(* IEC 61131-3 sources: daoli-st-library/DL_Algo (part 11) *)

(* ---- FB_DL_DewpointReset.st ---- *)
//==============================================================================
// 功能块：FB_DL_DewpointReset ｜ 中文名称：依据室内露点重置冷冻水供水温度设定
// 所属子库：DL_Algo ｜ 版本：v1.0.0 ｜ 兼容：CODESYS V3.5+ / TwinCAT 3 / 汇川 InoProShop
// 功能描述：室内露点重置冷冻水供水温度设定：目标 = max(露点 + 安全余
//           量, 下限)，带上下限钳位与斜率限制（fRateKPerS，由
//           uDeltaTimeMs 显式积分，禁系统时间函数）。露点由
//           FC_DL_DewPointCalc 计算（Magnus-Tetens 常数唯一属主为
//           FC_DL_VaporPressureSat，R23 裁定）——只调用不复制。双出
//           口：结露风险（露点 + 余量超上限，供水被顶到上限，除湿能
//           力不足，如实外显不静默）与域外钳位提示。失能保持设定。
// 开源溯源 (Origin)：道莅 clean-room 防御性实现（仅借 OSCAT ROOM_CONTROL 行为定义/参数域，零代码行与符号名复制）
// 单位表：温度[摄氏度] / 相对湿度[%] / 余量[K] / 斜率[K每s] / 扫描间隔[ms]
// 错误码表：16#0002_3601 信息级（露点域外钳位：湿度钳 1~100、干球钳
//           −40~60、下游件域外提示，不置 bError）/ 16#0002_3602 信息
//           级（防结露下限生效，供水被顶到上限，除湿能力不足，不置
//           bError）/ 16#0002_3605 预留禁用（不得挪用）/ 16#0002_3610
//           故障级（供水上下限倒置或余量/斜率组态非法，置 bError）/
//           16#0002_3611 故障级（输入非有限或下游件数据不可信，置
//           bError）/ 16#0002_3612 预留禁用（不得挪用）
// 状态机：E_DL_DewpointResetState（eIdle=0 / eTrack=10 / eCondRisk=20 /
//           eFault=99），CASE 含 ELSE 兜底，ELSE 复用 3611（§3 未为本
//           件单列兜底槽，不得越段加码）并回上限安全侧
// 边界行为：① 湿度钳 1~100、干球钳 −40~60（下游件承诺域），钳位发生
//           → 信息 3601；② 露点 + 余量大于供水上限 → bCondRisk :=
//           TRUE + 信息 3602，设定被顶到上限（如实反映「制冷量再低
//           也压不住露点」，不静默），退出条件两条：风险消失回追踪相
//           或失能回待机；③ fChwMinC 大于等于 fChwMaxC 或余量小于 0
//           或斜率非正 → 故障 3610；④ 非有限（NaN 自反判 + Inf 幅值
//           上限判，R79）→ 故障 3611，设定回供水上限安全侧（防结露
//           优先，冷却失效由上位温控回路告警，不静默）；⑤ 下游露点
//           件 uErrorId 非零或 bInRange 为假（预钳位后正常不可达，防
//           御路径）→ 复用信息 3601 且露点取干球温度保守估计（热力学
//           事实：露点不超过干球），下游信息级不升格（R115 纪律反向
//           适用：信息安全侧不得放大）；⑥ 失能 → 保持设定 + bValid :=
//           FALSE（供水温度突变会导致除湿振荡）；⑦ 斜率限制用
//           uDeltaTimeMs 显式积分，间隔为 0 本拍不动；⑧ 首拍设定从
//           下限起坡（首拍不出未知值）。
// 修订历史：v1.0.0 2026-11-17 首版（R25 派单 · §4.9）
//==============================================================================
(*------------------------------------------------------------------------------
 * 枚举: E_DL_DewpointResetState（归属 DL_Algo，与 FB_DL_DewpointReset 同文件）
 *----------------------------------------------------------------------------*)
TYPE E_DL_DewpointResetState :
(
    eIdle     := 0,   // 失能/待机：设定保持 / Idle: setpoint held
    eTrack    := 10,  // 斜率追踪：向目标设定限速逼近 / Track: rate-limited approach to target
    eCondRisk := 20,  // 结露风险：目标超上限，供水顶上限 / Condensation risk: target above ceiling, supply pinned
    eFault    := 99   // 故障兜底态：组态非法/非有限/非法状态，设定回上限 / Fault fallback, setpoint at ceiling
);
END_TYPE
FUNCTION_BLOCK FB_DL_DewpointReset
VAR_INPUT
    fRoomTempC    : LREAL;                     // 室内干球温度 [摄氏度] / Room dry-bulb temperature [degC]
    fRoomRhPct    : LREAL;                     // 室内相对湿度 [百分数] / Room relative humidity [percent]
    fChwMinC      : LREAL := 7.0;              // 供水设定下限 [摄氏度] / Chilled-water setpoint floor [degC]
    fChwMaxC      : LREAL := 18.0;             // 供水设定上限 [摄氏度] / Chilled-water setpoint ceiling [degC]
    fDewMarginK   : LREAL := 1.5;              // 防结露安全余量 [K] / Anti-condensation margin [K]
    fRateKPerS    : LREAL := 0.05;             // 设定斜率 [K每s] / Setpoint rate limit [K per s]
    uDeltaTimeMs  : UDINT;                     // 扫描间隔 [ms]，调用方注入，禁用系统时间函数 / Scan interval [ms], caller-injected
    bEnable       : BOOL;                      // 总使能 / Master enable
    bReset        : BOOL;                      // 复位，上升沿清状态与设定 / Reset, rising edge clears state and setpoint
END_VAR
VAR_OUTPUT
    fChwSetC      : LREAL;                     // 冷冻水供水温度设定 [摄氏度] / Chilled-water supply setpoint [degC]
    fDewPointC    : LREAL;                     // 室内露点 [摄氏度]，下游件计算透传 / Room dew point [degC], passed through
    fMarginK      : LREAL;                     // 当前供水设定相对露点裕量 [K] / Margin of setpoint over dew point [K]
    bCondRisk     : BOOL;                      // 露点超出可调范围，除湿能力不足 / Dew point beyond adjustable range, dehumidification short
    bAtMin        : BOOL;                      // 设定贴下限 / Setpoint at floor
    bAtMax        : BOOL;                      // 设定贴上限 / Setpoint at ceiling
    eErr          : UDINT;                     // 错误码，0 = 无错，码位 16#0002_3601 起信息级、16#0002_3610 起故障级（分带见错误码表） / Error code, 0 = no error, band info/fault per the code table
    bError        : BOOL;                      // 故障级标志，仅故障级错误置位 / Fault-class flag, set only on fault-level codes
    bValid        : BOOL;                      // 设定数据可用标志，失能/故障闸显式 FALSE / Setpoint usable flag, explicit FALSE on disable/fault gates
    eState        : E_DL_DewpointResetState;   // 主状态机当前状态 / Current state of the main state machine
END_VAR
VAR
    fbReset       : R_TRIG;                    // 复位上升沿检测实例 / Reset rising edge detector
    fRhClamped    : LREAL;                     // 钳位后湿度 [百分数] / Clamped humidity [percent]
    fTempClamped  : LREAL;                     // 钳位后干球 [摄氏度] / Clamped dry-bulb [degC]
    bDomainClamp  : BOOL;                      // 本拍发生域外钳位 / Domain clamp occurred this scan
    fTempReal     : REAL;                      // 干球降精度暂存 [摄氏度] / Dry-bulb staging in REAL precision
    fRhReal       : REAL;                      // 湿度降精度暂存 [百分数] / Humidity staging in REAL precision
    fDewReal      : REAL;                      // 露点返回值暂存 [摄氏度] / Dew-point return staging in REAL precision
    uDewErr       : UDINT;                     // 下游件错误码暂存 / Downstream error code staging
    fVaporPa      : REAL;                      // 下游件水汽压暂存 [Pa]（诊断透传）/ Downstream vapor pressure staging [Pa]
    bDewInRange   : BOOL;                      // 下游件域内标志暂存 / Downstream in-domain flag staging
    bDewOk        : BOOL;                      // 下游件结果可用判据 / Downstream result usable predicate
    fTargetC      : LREAL;                     // 钳位前目标设定 [摄氏度] / Pre-limit target setpoint [degC]
    fStepK        : LREAL;                     // 本拍允许步长 [K] / Allowed step this scan [K]
    fDeltaK       : LREAL;                     // 本拍目标增量 [K] / Target delta this scan [K]
    fDeltaApplied : LREAL;                     // 本拍实际增量 [K]（步长限幅后）/ Applied delta after rate limit [K]
    bFirstScan    : BOOL := TRUE;              // 首拍初始化标志 / First-scan initialization flag
END_VAR
VAR CONSTANT
    DL_DPR_CODE_INFO_1 : UDINT := 16#0002_3601;   // 信息级槽 1（露点域外钳位） / info slot 1
    DL_DPR_CODE_INFO_2 : UDINT := 16#0002_3602;   // 信息级槽 2（防结露下限生效） / info slot 2
    DL_DPR_CODE_RSV_1  : UDINT := 16#0002_3605;   // 预留禁用（不得挪用） / reserved, do not use
    DL_DPR_CODE_FLT_1  : UDINT := 16#0002_3610;   // 故障级槽 1（供水界倒置或组态非法） / fault slot 1
    DL_DPR_CODE_FLT_2  : UDINT := 16#0002_3611;   // 故障级槽 2（输入非有限） / fault slot 2
    DL_DPR_CODE_RSV_2  : UDINT := 16#0002_3612;   // 预留禁用（不得挪用） / reserved, do not use
    DL_DP_ZERO    : LREAL := 0.0;              // 零值常量，避免裸字面量 [—] / Zero constant, avoids a bare literal
    DL_DP_TOL     : LREAL := 1.0E-6;           // 浮点比较容差 [—] / Float comparison tolerance
    DL_DP_INF     : LREAL := 1.7976931348623157E308;  // LREAL 幅值上限，Inf 判据 / LREAL magnitude ceiling, Inf criterion
    DL_DP_RH_MIN  : LREAL := 1.0;              // 湿度钳位下限 [百分数] / Humidity clamp floor [percent]
    DL_DP_RH_MAX  : LREAL := 100.0;            // 湿度钳位上限 [百分数] / Humidity clamp ceiling [percent]
    DL_DP_T_MIN   : LREAL := -40.0;            // 干球钳位下限 [摄氏度]，下游件承诺域 / Dry-bulb clamp floor, downstream promised domain
    DL_DP_T_MAX   : LREAL := 60.0;             // 干球钳位上限 [摄氏度] / Dry-bulb clamp ceiling [degC]
    DL_DP_MS_PER_S : LREAL := 1000.0;          // 毫秒转秒系数 [s/ms] / Ms-to-s factor
END_VAR

(*------------------------------------------------------------------------------
 * 段 1｜无条件刷新区（红线 5）：复位沿检测在任何分支之外周期调用
 *----------------------------------------------------------------------------*)
fbReset(CLK := bReset);                        // 复位沿检测无条件刷新 / reset edge refreshed unconditionally

(*------------------------------------------------------------------------------
 * 段 2｜复位沿处理（改写置于沿后，防吞沿 R39）
 *----------------------------------------------------------------------------*)
IF fbReset.Q THEN
    eState  := E_DL_DewpointResetState.eIdle;
    eErr    := 16#0000_0000;                   // 复位清码 / reset clears code
    bError  := FALSE;                          // 复位清故障 / reset clears fault
    bCondRisk := FALSE;                        // 结露风险标志清 / condensation risk cleared
    bAtMin  := FALSE;                          // 贴下限清 / at-floor cleared
    bAtMax  := FALSE;                          // 贴上限清 / at-ceiling cleared
    bFirstScan := TRUE;                        // 重新首拍化 / re-initialize first scan
    fChwSetC := DL_DP_ZERO;                    // 设定清零待首拍初始化 / setpoint zeroed, awaits first-scan init
END_IF

(*------------------------------------------------------------------------------
 * 段 3｜非有限输入闸（浮点引脚逐个：NaN 自反判 + Inf 幅值上限判，R79）
 *       命中即设定回上限安全侧（防结露优先）
 *----------------------------------------------------------------------------*)
IF (fRoomTempC <> fRoomTempC) OR (ABS(fRoomTempC) >= DL_DP_INF)
   OR (fRoomRhPct <> fRoomRhPct) OR (ABS(fRoomRhPct) >= DL_DP_INF)
   OR (fChwMinC <> fChwMinC) OR (ABS(fChwMinC) >= DL_DP_INF)
   OR (fChwMaxC <> fChwMaxC) OR (ABS(fChwMaxC) >= DL_DP_INF)
   OR (fDewMarginK <> fDewMarginK) OR (ABS(fDewMarginK) >= DL_DP_INF)
   OR (fRateKPerS <> fRateKPerS) OR (ABS(fRateKPerS) >= DL_DP_INF) THEN
    eState  := E_DL_DewpointResetState.eFault;
    eErr    := DL_DPR_CODE_FLT_2;              // 故障级：输入非有限 / fault: non-finite input
    bError  := TRUE;                           // 故障级必置 bError（R45 配对）/ fault-class pairs with bError
    bValid  := FALSE;                          // 输出不可用 / outputs unusable
    fChwSetC := fChwMaxC;                      // 设定回上限安全侧（防结露优先）/ setpoint to ceiling, safe side
    bCondRisk := FALSE;                        // 故障态不判结露风险 / risk not judged in fault
    bAtMin := FALSE;                           // 贴限撤 / at-floor withdrawn
    bAtMax := TRUE;                            // 贴上限如实外显 / at-ceiling shown truthfully
    fDewPointC := DL_DP_ZERO;                  // 露点出口清零 / dew-point output zeroed
    fMarginK := DL_DP_ZERO;                    // 裕量出口清零 / margin output zeroed
    RETURN;
END_IF

(*------------------------------------------------------------------------------
 * 段 4｜组态合法性闸（供水界倒置/余量小于 0/斜率非正）
 *----------------------------------------------------------------------------*)
IF (fChwMinC >= fChwMaxC) OR (fDewMarginK < DL_DP_ZERO) OR (fRateKPerS <= DL_DP_TOL) THEN
    eState  := E_DL_DewpointResetState.eFault;
    eErr    := DL_DPR_CODE_FLT_1;              // 故障级：供水上下限倒置或组态非法 / fault: band inverted or config invalid
    bError  := TRUE;                           // 故障级必置 bError（R45 配对）/ fault-class pairs with bError
    bValid  := FALSE;                          // 输出不可用 / outputs unusable
    fChwSetC := fChwMaxC;                      // 设定回上限安全侧（防结露优先）/ setpoint to ceiling, safe side
    bCondRisk := FALSE;                        // 故障态不判结露风险 / risk not judged in fault
    bAtMin := FALSE;                           // 贴限撤 / at-floor withdrawn
    bAtMax := TRUE;                            // 贴上限如实外显 / at-ceiling shown truthfully
    fDewPointC := DL_DP_ZERO;                  // 露点出口清零 / dew-point output zeroed
    fMarginK := DL_DP_ZERO;                    // 裕量出口清零 / margin output zeroed
    RETURN;
END_IF

(*------------------------------------------------------------------------------
 * 段 5｜首拍初始化：设定从下限起坡（首拍不出未知值）
 *----------------------------------------------------------------------------*)
IF bFirstScan THEN
    fChwSetC := fChwMinC;                      // 首拍设定 = 下限 / first-scan setpoint = floor
    bFirstScan := FALSE;                       // 初始化完成 / initialization done
END_IF

(*------------------------------------------------------------------------------
 * 段 6｜域钳位（湿度 1~100、干球 −40~60，下游件承诺域）+ 露点组合调用
 *       （FC_DL_DewPointCalc，每拍恰好一次，只调用不复制）
 *----------------------------------------------------------------------------*)
fRhClamped := fRoomRhPct;                      // 湿度工作副本 / humidity working copy
fTempClamped := fRoomTempC;                    // 干球工作副本 / dry-bulb working copy
bDomainClamp := FALSE;                         // 钳位标志逐拍重判 / clamp flag re-judged per scan
IF fRhClamped < DL_DP_RH_MIN THEN
    fRhClamped := DL_DP_RH_MIN;                // 湿度钳下限 / humidity clamped to floor
    bDomainClamp := TRUE;                      // 钳位发生 / clamped
END_IF
IF fRhClamped > DL_DP_RH_MAX THEN
    fRhClamped := DL_DP_RH_MAX;                // 湿度钳上限 / humidity clamped to ceiling
    bDomainClamp := TRUE;                      // 钳位发生 / clamped
END_IF
IF fTempClamped < DL_DP_T_MIN THEN
    fTempClamped := DL_DP_T_MIN;               // 干球钳下限 / dry-bulb clamped to floor
    bDomainClamp := TRUE;                      // 钳位发生 / clamped
END_IF
IF fTempClamped > DL_DP_T_MAX THEN
    fTempClamped := DL_DP_T_MAX;               // 干球钳上限 / dry-bulb clamped to ceiling
    bDomainClamp := TRUE;                      // 钳位发生 / clamped
END_IF
fTempReal := LREAL_TO_REAL(fTempClamped);      // 干球降精度显式转换 / dry-bulb explicit narrowing
fRhReal := LREAL_TO_REAL(fRhClamped);          // 湿度降精度显式转换 / humidity explicit narrowing
fDewReal := FC_DL_DewPointCalc(fTempC := fTempReal, fRhPct := fRhReal,
                               uErrorId => uDewErr, fVaporPa => fVaporPa,
                               bInRange => bDewInRange);  // 露点组合调用，返回值即露点 [摄氏度] / dew-point call, return is the dew point
bDewOk := (uDewErr = 16#0000_0000) AND bDewInRange;    // 下游可用判据 / downstream usable predicate
IF bDewOk THEN
    fDewPointC := fDewReal;                    // 露点出口透传 / dew-point output pass-through
ELSE
    fDewPointC := fTempClamped;                // 防御路径：露点取干球保守估计（露点不超过干球）/ defensive: dry-bulb conservative estimate
    bDomainClamp := TRUE;                      // 下游域外提示并入钳位信息（不升格）/ downstream hint merged into clamp info
END_IF

(*------------------------------------------------------------------------------
 * 段 7｜目标计算：max(露点 + 余量, 下限)，超上限则顶上限并置结露风险
 *----------------------------------------------------------------------------*)
fTargetC := fDewPointC + fDewMarginK;          // 防结露目标 = 露点 + 余量 [摄氏度] / target = dew point plus margin
IF fTargetC < fChwMinC THEN
    fTargetC := fChwMinC;                      // 低于下限抬到下限 / below floor raised to floor
END_IF
IF fTargetC > fChwMaxC THEN
    fTargetC := fChwMaxC;                      // 超上限顶到上限 / above ceiling pinned to ceiling
END_IF

(*------------------------------------------------------------------------------
 * 段 8｜状态机：CASE 含 ELSE 兜底（非法状态 → 复用 3611 + 回上限，安全侧）
 *----------------------------------------------------------------------------*)
CASE eState OF

    E_DL_DewpointResetState.eIdle:
        bValid := FALSE;                       // 失能闸显式不可用（R72）/ explicit FALSE on disable gate
        bCondRisk := FALSE;                    // 待机不判风险 / risk not judged in idle
        bAtMin := FALSE;                       // 贴限撤 / at-floor withdrawn
        bAtMax := FALSE;                       // 贴限撤 / at-ceiling withdrawn
        eErr := 16#0000_0000;                  // 待机无错 / no error in idle
        bError := FALSE;                       // 待机无故障 / no fault in idle
        IF bEnable THEN
            eState := E_DL_DewpointResetState.eTrack;  // 使能进追踪相 / enable enters track
        END_IF

    E_DL_DewpointResetState.eTrack:
        bValid := TRUE;                        // 追踪相设定可用 / setpoint usable in track
        eErr := 16#0000_0000;                  // 追踪相先清码 / track clears code first
        bError := FALSE;                       // 追踪相先清故障 / track clears fault first
        IF bDomainClamp THEN
            eErr := DL_DPR_CODE_INFO_1;        // 信息级：露点域外钳位 / info: dew-point domain clamp
        END_IF
        IF NOT bEnable THEN
            eState := E_DL_DewpointResetState.eIdle;   // 失能回待机（设定保持）/ disable returns to idle, setpoint held
            bValid := FALSE;                   // 失能闸显式不可用 / explicit FALSE on disable gate
        ELSE
            fStepK := fRateKPerS * UDINT_TO_LREAL(uDeltaTimeMs) / DL_DP_MS_PER_S;  // 本拍步长 = 斜率乘时长 [K]，间隔 0 即不动 / step = rate times interval
            fDeltaK := fTargetC - fChwSetC;    // 目标增量 [K] / target delta [K]
            IF ABS(fDeltaK) <= fStepK THEN
                fDeltaApplied := fDeltaK;      // 一步到位 / single-step arrival
            ELSIF fDeltaK > DL_DP_ZERO THEN
                fDeltaApplied := fStepK;       // 正向限速 / positive rate-limited
            ELSE
                fDeltaApplied := -fStepK;      // 反向限速 / negative rate-limited
            END_IF
            fChwSetC := fChwSetC + fDeltaApplied;      // 限速逼近目标 / rate-limited approach
            bAtMin := ABS(fChwSetC - fChwMinC) < DL_DP_TOL;    // 贴下限（容差比较）/ at-floor with tolerance
            bAtMax := ABS(fChwSetC - fChwMaxC) < DL_DP_TOL;    // 贴上限（容差比较）/ at-ceiling with tolerance
            IF (fDewPointC + fDewMarginK) > fChwMaxC + DL_DP_TOL THEN
                eState := E_DL_DewpointResetState.eCondRisk;   // 露点超上限转结露风险相 / dew point beyond ceiling enters risk
            END_IF
        END_IF

    E_DL_DewpointResetState.eCondRisk:
        bValid := TRUE;                        // 风险相设定可用（顶上限值）/ setpoint usable in risk (pinned value)
        fChwSetC := fChwMaxC;                  // 供水被顶到上限（除湿能力不足，如实外显）/ supply pinned to ceiling
        bCondRisk := TRUE;                     // 结露风险标志 / condensation risk flag
        bAtMin := FALSE;                       // 贴下限撤 / at-floor withdrawn
        bAtMax := TRUE;                        // 贴上限如实外显 / at-ceiling shown truthfully
        eErr := DL_DPR_CODE_INFO_2;            // 信息级：防结露下限生效 / info: anti-condensation limit active
        bError := FALSE;                       // 信息级不置 bError / info never raises bError
        IF NOT bEnable THEN
            eState := E_DL_DewpointResetState.eIdle;   // 失能回待机（第二条退出条件）/ disable returns to idle, second exit
            bValid := FALSE;                   // 失能闸显式不可用 / explicit FALSE on disable gate
            bCondRisk := FALSE;                // 风险标志清 / risk flag cleared
        ELSIF (fDewPointC + fDewMarginK) <= fChwMaxC + DL_DP_TOL THEN
            eState := E_DL_DewpointResetState.eTrack;  // 风险消失回追踪相（第一条退出条件）/ risk gone, first exit to track
        END_IF

    ELSE
        eState := E_DL_DewpointResetState.eFault;  // 非法状态兜底 / illegal-state fallback
        eErr := DL_DPR_CODE_FLT_2;             // 兜底复用故障级槽 2（§3 未单列兜底槽，不得越段加码）/ fallback reuses fault slot 2
        bError := TRUE;                        // 故障级必置 bError / fault-class pairs with bError
        bValid := FALSE;                       // 输出不可用 / outputs unusable
        fChwSetC := fChwMaxC;                  // 设定回上限安全侧（防结露优先）/ setpoint to ceiling, safe side
        bCondRisk := FALSE;                    // 风险标志清 / risk flag cleared
        bAtMin := FALSE;                       // 贴限撤 / at-floor withdrawn
        bAtMax := TRUE;                        // 贴上限如实外显 / at-ceiling shown truthfully
END_CASE

(*------------------------------------------------------------------------------
 * 段 9｜裕量出口：当前供水设定相对露点裕量 [K]（负值即结露，可观测）
 *----------------------------------------------------------------------------*)
fMarginK := fChwSetC - fDewPointC;             // 裕量 = 设定 − 露点 [K] / margin = setpoint minus dew point
END_FUNCTION_BLOCK

(* ---- FB_DL_Differentiator.st ---- *)
(*==============================================================================
 * 组件名称 (Component)  : FB_DL_Differentiator
 * 所属子库 (Sublibrary) : DL_Algo
 * 当前版本 (Version)    : 1.0.1
 * 兼容性   (Platform)   : CODESYS 3.5 / TwinCAT 3 / 汇川 InoProShop / Machine Expert
 *                         仅依赖 Standard.library（LIMIT / MIN / MAX / ABS），零厂商方言
 * 功能描述 (Function)   : 带一阶低通滤波的实用微分器：差分商 (fIn - fInPrev)/fDt
 *                         计算变化率，后接一阶低通抑制高频噪声放大（纯差分对
 *                         采样噪声增益 1/fDt，会放大毛刺）。输出变化率限幅
 *                         （rRateMin/rRateMax）防异常尖峰误触发趋势报警。
 *                         现场用途：温度变化速率监控（趋势报警前级）、压装
 *                         速度计算、液位升降速率。
 * 开源溯源 (Origin)     : 原创实现。组合语义对应西门子 LGF 的差分商块与
 *                         PT1 滤波器串联的公开行为定义，clean-room 编写，
 *                         未复制任何厂商私有库源码。
 * 本文件内含       : TYPE  E_DL_DiffState（配套枚举，归属 DL_Algo）
 *                    FB    FB_DL_Differentiator
 * 依赖     (Depends)    : 无 DL_ 内部依赖；Standard.library: LIMIT / MIN / MAX / ABS
 * 红线自检 (Redline)    : R1 ✓ 零全局变量表与外部变量引用 ｜ R2 ✓ 零物理 IO 地址直写
 *                         R3 ✓ 纯 IEC 61131-3 ｜ R4 ✓ 防除零+钳位+非有限值拒绝
 *                         R5 ✓ 全变量中英双语同行注释 ｜ R6 ✓ 四态 ENUM+CASE+ELSE
 *                         R7 N/A（无定时器/边沿实例）
 * 【边界披露 / Boundary disclosure】
 *   B1 除零防御：fDt 走公共钳位（<10ms 钳位 10ms 置 16#0002_0002），恒大于零。
 *   B2 tFiltTime 超上限 60s：钳位并置 16#0002_1401；tFiltTime=0 为合法直通
 *      （输出原始差分商，不置故障）。
 *   B3 rRateMin > rRateMax：自动对调并置 16#0002_0001。
 *   B4 输入非有限值：本拍拒绝、清历史（bHistValid=FALSE）、输出归零，置
 *      16#0002_0004；下一有效拍重新同步端点，绝不输出伪造速率。
 *   B5 首扫同步 fInPrev := fIn、输出 0，防上电尖峰。
 *   B6 低通系数 fAlpha 显式钳位 0..1；fTfEff + fDt 恒 > 0（分母安全）。
 * 【验收向量 / Acceptance vectors】
 *   V1  fIn 每拍 +1.0（tSampleTime=100MS，即 10 EU/s 恒速）→ fRawRate=10 EU/s，
 *       fRateOut 数拍内收敛到 10 EU/s、bValid=TRUE
 *   V2  fIn 阶跃 +50 一拍 → fRawRate=500 EU/s 单拍尖峰，fRateOut 按
 *       tFiltTime=500MS 平滑，峰值明显低于 500（噪声抑制效果）
 *   V3  fIn 恒定 → fRateOut 收敛到 0
 *   V4  rRateMax=20，V1 → fRateOut 钳位 20 EU/s
 *   V5  tFiltTime=0 → fRateOut=fRawRate（直通，无故障码）
 *   V6  tFiltTime=65S → 钳位 60S、16#0002_1401
 *   V7  fIn=NaN → 16#0002_0004，fRateOut=0、bValid=FALSE
 * 修订历史 (Revision)   :
 *   2026-11-15  v1.0.0  首版入库（Round 04 · Phase 3 · DL_Algo 批次）
 *   2026-11-15  v1.0.1  阶段五终审精修：首扫初始化标志判据修复（原判据恒假
 *                       为死代码），首扫同步端点改为显式可审计路径
 *============================================================================*)

(*-----------------------------------------------------------------------------
 * 枚举: E_DL_DiffState（归属 DL_Algo，与 FB_DL_Differentiator 同文件）
 * 含义: 微分器状态机离散状态。数值步长留空位便于后续插态而不破坏已有工程。
 *----------------------------------------------------------------------------*)
TYPE E_DL_DiffState :
(
    eInit  := 0,   // 初始化态：首扫或失历史，同步端点、输出清零 / Init state, sync endpoint, output zero
    eRun   := 10,  // 运行态：差分商 + 低通滤波逐拍计算 / Run state, difference quotient with low-pass per scan
    eTrack := 20,  // 跟踪态：输出立即跟随 fTrackValue / Track state, output follows track value instantly
    eFault := 99   // 故障兜底态：非法状态拦截，自动回初始化 / Fault fallback, auto recover to init
);
END_TYPE

(*==============================================================================
 * 功能块: FB_DL_Differentiator
 * 调用约定: 每个扫描周期无条件调用一次；bTrack 使能时输出立即跟随 fTrackValue。
 * 无状态泄漏: 全部状态驻留于实例私有 VAR，可多实例并行互不影响。
 * 噪声披露: 输出滞后 ≈ tFiltTime；tFiltTime 越小噪声抑制越弱，建议
 *           tFiltTime >= 5 × 采样周期（本块默认 500ms @ 100ms 采样）。
 *============================================================================*)
FUNCTION_BLOCK FB_DL_Differentiator
VAR_INPUT
    bEnable     : BOOL := FALSE;      // 使能标志，FALSE 时输出 0 / Enable flag, FALSE forces output to zero
    fIn         : REAL := 0.0;        // 被微分量 [EU]，如温度/位置/液位 / Differentiated input [EU]
    tFiltTime   : TIME := T#500MS;    // 速率低通时间常数 [s]，0 = 原始差分直通 / Rate low-pass time constant [s], 0 = raw pass
    rRateMin    : REAL := -1.0E10;    // 速率下限 [EU/s]，大于上限时自动对调 / Rate lower limit [EU/s], swapped if greater
    rRateMax    : REAL := 1.0E10;     // 速率上限 [EU/s]，小于下限时自动对调 / Rate upper limit [EU/s], swapped if smaller
    bTrack      : BOOL := FALSE;      // 跟踪使能，TRUE 时输出立即跟随 fTrackValue / Track enable, output follows track value
    fTrackValue : REAL := 0.0;        // 跟踪值 [EU/s]，投切无扰动基准 / Track value [EU/s], bumpless transfer reference
    tSampleTime : TIME := T#100MS;    // 采样周期 [s]，小于 10ms 钳位为 10ms / Sample time [s], clamped to 10ms
END_VAR
VAR_OUTPUT
    fRateOut    : REAL;               // 变化率输出 [EU/s]，滤波并限幅 / Rate output [EU/s], filtered and limited
    fRawRate    : REAL;               // 未滤波原始速率 [EU/s]，诊断 / Raw unfiltered rate [EU/s] for diagnostics
    bValid      : BOOL;               // 输出有效标志（端点已同步且有真实差分）/ Output valid flag
    bError      : BOOL;               // 故障标志（瞬时，逐拍重算） / Fault flag, transient, recomputed every scan
    uErrorId    : UDINT;              // 故障码，0 = 无故障 / Error code, 0 = no error
END_VAR
VAR
    fInPrev     : REAL;               // 上一拍被微分量 [EU]，差分端点 / Previous input [EU], difference endpoint
    fTfEff      : REAL;               // 钳位后滤波时间常数 [s] / Clamped filter time constant [s]
    fAlpha      : REAL;               // 低通滤波系数 [0..1] / Low-pass filter coefficient [0..1]
    fDt         : REAL;               // 折算后的采样周期 [s] / Converted sample period [s]
    bInFinite   : BOOL;               // 本拍输入有限值标志 / Input finite validity flag this scan
    bHistValid  : BOOL;               // 端点历史有效标志 / Endpoint history valid flag
    bInit       : BOOL;               // 首扫标志 / First scan flag
    eState      : E_DL_DiffState;     // 主状态机当前状态 / Current state of the main state machine
END_VAR
VAR CONSTANT
    DL_DIFF_TF_MAX : REAL := 60.0;    // 滤波时间常数上限 [s] / Filter time constant upper limit [s]
    DL_DIFF_EPS    : REAL := 1.0E-6;  // 分母安全容差 / Denominator safety tolerance
END_VAR

(*------------------------------------------------------------------------------
 * 段 1｜公共参数处理（通用约定 0-1/0-2/0-3）：周期钳位、滤波常数钳位、量程对调
 *      Common handling: sample time clamp, filter constant clamp, limit swap
 *-----------------------------------------------------------------------------*)
uErrorId := 16#0000_0000;               // 故障码逐拍重算 / Error code recomputed every scan
bError   := FALSE;                      // 故障标志逐拍重算 / Fault flag recomputed every scan

IF tSampleTime < T#10MS THEN
    fDt      := TIME_TO_REAL(T#10MS) / 1000.0; // 非法周期钳位为 10ms（边界 B1 防除零）/ Illegal period clamped to 10ms
    uErrorId := 16#0002_0002;           // 采样周期非法已钳位 / Sample time illegal, clamped
ELSE
    fDt      := TIME_TO_REAL(tSampleTime) / 1000.0; // 周期换算为秒 [s] / Period converted to seconds [s]
END_IF

fTfEff := TIME_TO_REAL(tFiltTime) / 1000.0; // 滤波常数换算为秒 [s] / Filter constant converted to seconds [s]
IF fTfEff < 0.0 THEN
    fTfEff   := 0.0;                    // 负值钳位为直通 / Negative clamped to pass-through
    uErrorId := 16#0002_1401;           // 滤波时间常数非法已钳位 / Filter time constant illegal, clamped
END_IF
IF fTfEff > DL_DIFF_TF_MAX THEN
    fTfEff   := DL_DIFF_TF_MAX;         // 超上限钳位（边界 B2）/ Over-limit clamped
    uErrorId := 16#0002_1401;           // 滤波时间常数非法已钳位 / Filter time constant illegal, clamped
END_IF

IF rRateMin > rRateMax THEN
    rRateMin := rRateMin + rRateMax;    // 三步对调第一步：求和 / Swap step one: sum
    rRateMax := rRateMin - rRateMax;    // 三步对调第二步：得旧下限 / Swap step two: old lower limit
    rRateMin := rRateMin - rRateMax;    // 三步对调第三步：得旧上限 / Swap step three: old upper limit
    uErrorId := 16#0002_0001;           // 参数越界已对调 / Limits out of order, swapped
END_IF

(*------------------------------------------------------------------------------
 * 段 2｜输入合法性（边界 B4）：非有限值拒绝并清历史，输出归零防伪造速率
 *      Input validity: non-finite rejected, history cleared, output zeroed
 *-----------------------------------------------------------------------------*)
bInFinite := NOT (fIn <> fIn) AND (ABS(fIn) <= 1.0E30); // NaN 判别 + 幅值防御 / NaN check plus magnitude guard

IF NOT bInFinite THEN
    uErrorId   := 16#0002_0004;         // 输入非有限值已拒绝 / Non-finite input rejected
    bHistValid := FALSE;                // 清历史端点 / Clear endpoint history
    fRateOut   := 0.0;                  // 输出归零 / Output zeroed
    fRawRate   := 0.0;                  // 原始速率归零 / Raw rate zeroed
    bValid     := FALSE;                // 有效标志清零 / Valid flag cleared
    eState     := eInit;                // 回初始化态重新同步 / Back to init for re-sync
END_IF

(*------------------------------------------------------------------------------
 * 段 3｜跟踪与首扫（约定 0-6）：端点同步、输出归零，防上电尖峰（边界 B5）
 *      Tracking and first scan: endpoint synced, output zeroed against power-up spike
 *-----------------------------------------------------------------------------*)
IF NOT bInit THEN
    IF bInFinite THEN
        fInPrev := fIn;                 // 端点同步当前输入 / Endpoint synced to current input
        bHistValid := TRUE;             // 历史有效 / History valid
    END_IF
    fRateOut := 0.0;                    // 输出清零 / Output zeroed
    fRawRate := 0.0;                    // 原始速率清零 / Raw rate zeroed
    bValid   := FALSE;                  // 首扫无真实差分 / No real difference on first scan
    eState   := eInit;                  // 回初始化态 / Back to init state
    bInit    := TRUE;                   // 首扫标志置位 / First scan flag set
END_IF

IF bTrack THEN
    fRateOut := LIMIT(rRateMin, fTrackValue, rRateMax); // 输出立即跟随跟踪值并限幅 / Output follows track value with limits
    IF bInFinite THEN
        fInPrev := fIn;                 // 端点同步当前输入 / Endpoint synced to current input
    END_IF
    bHistValid := TRUE;                 // 历史有效 / History valid
    bValid     := TRUE;                 // 跟踪输出视为有效 / Tracked output considered valid
    eState     := eTrack;               // 跟踪态 / Track state
END_IF

(*------------------------------------------------------------------------------
 * 段 4｜使能失效语义：输出归零、清历史，恢复后从初始化态重新同步
 *      Disabled semantics: output zeroed, history cleared, re-sync after enable
 *-----------------------------------------------------------------------------*)
IF NOT bEnable THEN
    fRateOut   := 0.0;                  // 输出归零 / Output zeroed
    fRawRate   := 0.0;                  // 原始速率归零 / Raw rate zeroed
    bValid     := FALSE;                // 有效标志清零 / Valid flag cleared
    bHistValid := FALSE;                // 清历史端点 / Clear endpoint history
    eState     := eInit;                // 回初始化态 / Back to init state
ELSE
    (*--------------------------------------------------------------------------
     * 段 5｜主状态机（红线 R6）：四态 ENUM + CASE + ELSE 兜底
     *     Main state machine: four-state ENUM + CASE with mandatory ELSE fallback
     *-------------------------------------------------------------------------*)
    CASE eState OF

        eInit:  // 初始化态：端点同步、输出 0，下拍进入运行态（边界 B5）/ Init: sync endpoint, output zero
            IF bInFinite THEN
                fInPrev := fIn;             // 端点同步当前输入 / Endpoint synced to current input
                bHistValid := TRUE;         // 历史有效 / History valid
            END_IF
            fRateOut := 0.0;                // 输出清零 / Output zeroed
            fRawRate := 0.0;                // 原始速率清零 / Raw rate zeroed
            bValid   := FALSE;              // 本拍无真实差分 / No real difference this scan
            eState   := eRun;               // 进入运行态 / Enter run state

        eRun:  // 运行态：差分商 + 低通滤波（边界 B1 分母安全）/ Run: difference quotient with low-pass
            IF NOT bHistValid THEN
                fInPrev := fIn;             // 历史失效先重建端点 / Rebuild endpoint when history invalid
                bHistValid := TRUE;         // 历史恢复有效 / History restored
                fRateOut := 0.0;            // 输出先归零防尖峰 / Output zeroed against spike
                fRawRate := 0.0;            // 原始速率归零 / Raw rate zeroed
            ELSE
                fRawRate := (fIn - fInPrev) / fDt; // 原始差分商 [EU/s] / Raw difference quotient [EU/s]
                IF fTfEff <= DL_DIFF_EPS THEN
                    fAlpha := 1.0;          // 零滤波常数直通（边界 B2 合法）/ Zero constant pass-through
                ELSE
                    fAlpha := fDt / (fTfEff + fDt); // 一阶低通系数 [0..1] / First-order low-pass coefficient
                    fAlpha := MIN(MAX(fAlpha, 0.0), 1.0); // 系数显式钳位（边界 B6）/ Coefficient explicitly clamped
                END_IF
                fRateOut := fRateOut + fAlpha * (fRawRate - fRateOut); // 低通递推 [EU/s] / Low-pass recursion [EU/s]
                fRateOut := LIMIT(rRateMin, fRateOut, rRateMax); // 速率限幅 / Rate limited
                fInPrev  := fIn;            // 端点更新 / Endpoint updated
                bValid   := TRUE;           // 输出有效 / Output valid
            END_IF

        eTrack:  // 跟踪态：输出已由段 3 跟随，释放后回运行态 / Track: output follows, resume run after release
            IF NOT bTrack THEN
                eState := eRun;             // 释放跟踪，恢复计算 / Tracking released, resume computing
            END_IF

        eFault:  // 故障兜底态：输出归零并回初始化态（无锁死）/ Fault fallback: output zeroed, recover to init
            fRateOut := 0.0;                // 输出归零 / Output zeroed
            eState   := eInit;              // 自动恢复初始化 / Auto recover to init

        ELSE  // 非法状态拦截：任何未定义状态一律进故障态并置码 / Illegal state interception
            eState   := eFault;             // 强制故障态 / Force fault state
            uErrorId := 16#0002_0005;       // 非法状态兜底 / Illegal state fallback
            bError   := TRUE;               // 故障标志置位 / Fault flag set

    END_CASE;
END_IF
END_FUNCTION_BLOCK

(* ---- FB_DL_DisturbanceObserver.st ---- *)
(*
  FB_DL_DisturbanceObserver  —  模型法负载扰动观测器 / Model-based load disturbance observer
  分类 Category : DL_Algo
  码位 Code     : 16#02_3_81
  版本 Version  : 1.0.0
  来源标签 Tag  : t2-4-s7-motion
  溯源 Source   : S7 Motion Control 语义借鉴 · clean-room 实现，仅借分类/参数域/命名，未复制源码行
  功能 Function : 1) 标称模型逆（J·dω/dt ÷ Kt）折算等效电流，与指令电流之差乘 Kt 得扰动转矩估计；
                  2) 估计量经一阶 Q 滤波（委托 FB_DL_LowPassFilter）去噪后输出；
                  3) 补偿量按 fCompGain 加权并限幅到 ±fCompLimit，饱和置 bSaturated。
  边界 Boundary : ① fInertia / fTorqueConst / fQFilterTau / fRatedCurrentA 任一 <= 0 判组态错置码且不投运（防除零）；
                  ② 速度为零并持续超冻结窗 tZeroSpeedHold（本件常量 200 ms）时冻结估计（静止段无可观测加速度，防噪声灌入）；
                  ③ bEnable 下降沿清估计值与微分状态（R28-1 解除式 = bEnable 上升沿 + bReset，两路径均在引脚可满足）；
                  ④ 补偿限幅 fCompLimit 由引脚给出，不在本件硬编码；
                  ⑤ bEnable = FALSE 语义：输出降级为安全值 0 + 保持状态 eIdle，不冻结末值（R191 显式声明）。
  依赖 Depends  : FB_DL_LowPassFilter × 1（Q 滤波，每拍无条件调用）
  同拍双窗配比  : 冻结窗 tZeroSpeedHold = 200 ms 与 Q 滤波时间常数 fQFilterTau 同源于 fSampleDt；
                  配比约束 fQFilterTau <= 0.5 × tZeroSpeedHold 保证静止冻结前滤波器已收敛（R100）

  码表 Error codes（本件格 02_3_81，子码步进 +0x10）:
    16#0002_0281 故障级：组态非法（惯量 / 转矩常数 / 滤波时间常数 / 额定电流 <= 0，或采样周期 <= 0，或组态量非有限）
    16#0002_0291 故障级：相 ID 越界（枚举兜底路径，复用组态码段之外的单列码）
    16#0002_02A1 信息级：速度为零冻结估计 / 输入非有限本拍不更新（不置 bError）

  修订历史 Revision :
    2026-11-18  v1.0.0  R36 首版入库
*)

TYPE E_DL_ObserverState :
(
    eIdle  := 0,   // 空闲（未使能，输出降级为 0）/ Idle, outputs degraded to zero
    eRun   := 10,  // 观测运行 / Observer running
    eHold  := 20,  // 静止冻结（速度为零超冻结窗）/ Frozen at zero speed
    eFault := 90   // 组态故障锁定（需 bReset 沿解除）/ Configuration fault locked
);
END_TYPE

FUNCTION_BLOCK FB_DL_DisturbanceObserver
VAR_INPUT
    bEnable        : BOOL := FALSE;              // 总使能，FALSE 时输出降级为 0 并回 eIdle / Master enable
    bReset         : BOOL := FALSE;              // 复位，上升沿清组态故障锁存 / Reset, clears latched fault
    fCmdOut        : REAL := 0.0;                // 控制器输出（力矩指令）[% 额定力矩] / Controller output [% rated torque]
    fRatedCurrentA : REAL := 10.0;               // 额定电流 [A]，域 > 0 / Rated current [A], domain > 0
    fMeasSpeed     : REAL := 0.0;                // 实测转速 [rpm]，带符号 / Measured speed [rpm]
    fInertia       : REAL := 0.001;              // 折算惯量 [kg·m²]，域 > 0 / Reflected inertia [kg·m²]
    fTorqueConst   : REAL := 1.0;                // 转矩常数 [N·m/A]，域 > 0 / Torque constant [N·m/A]
    fQFilterTau    : REAL := 0.005;              // Q 滤波时间常数 [s]，域 > 0 / Q-filter time constant [s]
    tSampleTime    : TIME := T#10MS;             // 采样周期 [ms 口径]，域 > 0 / Sampling period
    fCompGain      : REAL := 1.0;                // 补偿加权系数 [1]，域 >= 0 / Compensation gain
    fCompLimitPct  : REAL := 20.0;               // 补偿限幅 [%]，域 > 0 / Compensation limit [%]
    fEps           : REAL := 1.0E-6;             // 浮点判零容差 [1] / Floating zero tolerance
END_VAR
VAR_OUTPUT
    fDistTorqueEst : REAL;                       // 扰动转矩估计 [N·m] / Estimated disturbance torque [N·m]
    fCompOut       : REAL;                       // 补偿量输出 [%]，限幅后 / Compensation output [%]
    bSaturated     : BOOL;                       // 补偿限幅饱和标志（单拍）/ Compensation saturated, single scan
    bFrozen        : BOOL;                       // 静止冻结标志 / Frozen at zero speed
    bValid         : BOOL;                       // 估计有效标志（单拍）/ Estimate valid, single scan
    bError         : BOOL;                       // 故障标志，派生自锁存 / Fault flag derived from latch
    uErrorId       : UDINT;                      // 事件码，0 = 无事件 / Event code, 0 = no event
    eStateOut      : E_DL_ObserverState;         // 状态出口，段尾单点映射 / State mapped at tail
END_VAR
VAR
    fbQFilter      : FB_DL_LowPassFilter;        // Q 滤波实例（每拍无条件调用）/ Q-filter instance
    tonZeroSpeed   : TON;                        // 零速持续时间窗（本件常量 200 ms）/ Zero-speed dwell timer
    rtEnable       : R_TRIG;                     // 使能上升沿 / Enable rising edge
    rtReset        : R_TRIG;                     // 复位上升沿 / Reset rising edge
    _eState        : E_DL_ObserverState := E_DL_ObserverState.eIdle;  // 内部状态机当前态 / Internal phase
    _uFault        : UDINT;                      // 故障码锁存（仅复位沿清除）/ Latched fault code
    _uInfo         : UDINT;                      // 信息码，每拍重算 / Information code, recomputed each scan
    _bFault        : BOOL;                       // 故障锁存位 / Latched fault bit
    fSpeedPrev     : REAL;                       // 上一拍转速快照 [rpm]（不参与预清零）/ Speed snapshot, kept
    fAccelRpmS     : REAL;                       // 转速微分 [rpm/s] / Speed derivative [rpm/s]
    fAccelRadS     : REAL;                       // 角加速度 [rad/s²] / Angular acceleration [rad/s²]
    fCurrentNomA   : REAL;                       // 标称模型逆等效电流 [A] / Nominal model inverse current [A]
    fCurrentCmdA   : REAL;                       // 指令折算电流 [A] / Command current [A]
    fTorqueDistNm  : REAL;                       // 含噪扰动转矩 [N·m] / Raw disturbance torque [N·m]
    fDtSec         : REAL;                       // 采样周期秒值 [s] / Sampling period in seconds
    bFirstScan     : BOOL := TRUE;               // 首扫标志（微分初值用）/ First-scan flag for derivative
    bZeroSpeed     : BOOL;                       // 零速判定中间量 / Zero-speed predicate
    bCfgBad        : BOOL;                       // 组态非法聚合标志 / Configuration invalid aggregate
END_VAR
VAR CONSTANT
    DL_T_ZERO_HOLD : TIME  := T#200MS;   // 零速冻结窗 [ms]，本件声明常量 / Zero-speed freeze window
    DL_RPM2RAD     : REAL  := 0.1047197551;  // rpm 转 rad/s [rad/(s·rpm)] / rpm to rad/s factor
    DL_EPS         : REAL  := 1.0E-6;    // 判零容差 [1] / Zero tolerance
END_VAR

(* —— 段 0：定时器与边缘检测无条件周期刷新（禁置于分支内） —— *)
rtEnable(CLK := bEnable);                                      // 使能上升沿（每拍必调）
rtReset(CLK := bReset);                                        // 复位上升沿（每拍必调）
bZeroSpeed := bEnable AND (ABS(fMeasSpeed) < DL_EPS);          // 零速判定，门控挂状态量
tonZeroSpeed(IN := bZeroSpeed, PT := DL_T_ZERO_HOLD);          // 零速驻留计时（输入非字面 TRUE，具备复位路径）

(* —— 段 1：单拍标志预清零（只清单拍量，快照与锁存不入清单） —— *)
bSaturated := FALSE;      // 单拍标志：限幅饱和
bValid     := FALSE;      // 单拍标志：估计有效
bFrozen    := FALSE;      // 单拍标志：静止冻结
bError     := FALSE;      // 单拍标志：故障出口（段 6 由锁存派生重写）
_uInfo     := 0;          // 信息码每拍重算
fDtSec     := TIME_TO_REAL(tSampleTime) / 1000.0;   // 采样周期秒值 [s]

(* —— 段 2：复位沿清故障锁存（R188 可达清除路径） —— *)
IF rtReset.Q THEN
    _bFault := FALSE;     // 复位沿清锁存位
    _uFault := 0;         // 复位沿清锁存码
END_IF

(* —— 段 3：组态域闸（覆盖全部参与换算的引脚，R151） —— *)
bCfgBad := FALSE;
IF (fInertia <> fInertia) OR (fInertia <= 0.0) THEN
    bCfgBad := TRUE;      // 惯量非有限或 <= 0
END_IF
IF (fTorqueConst <> fTorqueConst) OR (fTorqueConst <= 0.0) THEN
    bCfgBad := TRUE;      // 转矩常数非有限或 <= 0
END_IF
IF (fQFilterTau <> fQFilterTau) OR (fQFilterTau <= 0.0) THEN
    bCfgBad := TRUE;      // 滤波时间常数非有限或 <= 0
END_IF
IF (fRatedCurrentA <> fRatedCurrentA) OR (fRatedCurrentA <= 0.0) THEN
    bCfgBad := TRUE;      // 额定电流非有限或 <= 0
END_IF
IF (fCompLimitPct <> fCompLimitPct) OR (fCompLimitPct <= 0.0) THEN
    bCfgBad := TRUE;      // 补偿限幅非有限或 <= 0
END_IF
IF (fEps <> fEps) OR (fEps <= 0.0) THEN
    bCfgBad := TRUE;      // 判零容差非有限或 <= 0
END_IF
IF tSampleTime <= T#0MS THEN
    bCfgBad := TRUE;      // 采样周期 <= 0（微分除零前置）
END_IF
IF bCfgBad THEN
    _uFault := 16#0002_0281;                              // 故障级：组态非法
    _bFault := TRUE;                                      // 锁存位置位（复位沿可清）
    bError := TRUE;                                       // 故障标志置位（R45 配对）
    _eState := E_DL_ObserverState.eFault;                 // 状态机进故障相
END_IF

(* —— 段 4：观测内核（仅无故障且使能时执行） —— *)
IF (NOT _bFault) AND bEnable AND (fDtSec > 0.0) THEN
    fCurrentCmdA := fCmdOut / 100.0 * fRatedCurrentA;                    // 指令折算电流 [A]
    IF bFirstScan THEN
        fSpeedPrev := fMeasSpeed;                                        // 首扫微分初值，防冲击
        bFirstScan := FALSE;                                             // 首扫标志唯一置假点
    END_IF
    fAccelRpmS := (fMeasSpeed - fSpeedPrev) / fDtSec;                    // 转速微分 [rpm/s]
    fAccelRadS := fAccelRpmS * DL_RPM2RAD;                               // 角加速度 [rad/s²]
    fSpeedPrev := fMeasSpeed;                                            // 快照更新（末行，不预清零）
    fCurrentNomA := fInertia * fAccelRadS / fTorqueConst;                // 标称模型逆等效电流 [A]（Kt 已证 > 0）
    fTorqueDistNm := (fCurrentCmdA - fCurrentNomA) * fTorqueConst;       // 含噪扰动转矩 [N·m]
    IF tonZeroSpeed.Q THEN
        _eState := E_DL_ObserverState.eHold;                             // 静止冻结相
        bFrozen    := TRUE;                                                // 冻结标志（出口 bFrozen，VAR_OUTPUT）
        _uInfo := 16#0002_02A1;                                         // 信息级：速度为零冻结估计
    ELSE
        _eState := E_DL_ObserverState.eRun;                             // 观测运行相
        fbQFilter(bEnable := TRUE, fIn := fTorqueDistNm, tTimeConst := REAL_TO_TIME(fQFilterTau * 1000.0),
                  tSampleTime := tSampleTime);                          // Q 滤波实例调用（每拍必调，单点单次）
        IF fbQFilter.bError THEN
            _eState := E_DL_ObserverState.eHold;                        // 滤波故障降级为冻结（降级不抛故障，R191 已声明）
        END_IF
    END_IF
ELSE
    _eState := E_DL_ObserverState.eIdle;                                // 未使能：降级为安全值（R191 声明）
    fSpeedPrev := fMeasSpeed;                                           // 快照跟随，防再使能冲击
    bFirstScan := TRUE;                                                 // 复位首扫标志（再使能重新取值）
END_IF

(* —— 段 5：状态机兜底（非法枚举值回 eIdle 并置故障级码） —— *)
CASE _eState OF
E_DL_ObserverState.eIdle:
    fCompOut := 0.0;                     // 空闲：补偿量降级为 0
    fDistTorqueEst := 0.0;               // 空闲：估计值清零
E_DL_ObserverState.eRun:
    fDistTorqueEst := fbQFilter.fOut;    // 运行：输出滤波后扰动估计 [N·m]
    fCompOut := -fCompGain * fDistTorqueEst / fTorqueConst / fRatedCurrentA * 100.0;  // 补偿量 [%]（Kt、额定电流已证 > 0）
    IF fCompOut > fCompLimitPct THEN
        fCompOut := fCompLimitPct;       // 上行限幅
        bSaturated := TRUE;              // 饱和标志
    ELSIF fCompOut < -fCompLimitPct THEN
        fCompOut := -fCompLimitPct;      // 下行限幅
        bSaturated := TRUE;              // 饱和标志
    END_IF
    bValid := TRUE;                      // 本拍估计有效
E_DL_ObserverState.eHold:
    fDistTorqueEst := 0.0;               // 冻结：不出新估计（静止段无可观测加速度）
    fCompOut := 0.0;                     // 冻结：补偿量 0
E_DL_ObserverState.eFault:
    fDistTorqueEst := 0.0;               // 故障：输出安全值
    fCompOut := 0.0;                     // 故障：输出安全值
ELSE
    _uFault := 16#0002_0291;             // 故障级：相 ID 越界（枚举兜底）
    _bFault := TRUE;                     // 锁存位置位
    bError := TRUE;                      // 故障标志置位（R45 配对）
    _eState := E_DL_ObserverState.eFault;  // 强制回故障相
    fDistTorqueEst := 0.0;               // 兜底输出安全值
    fCompOut := 0.0;                     // 兜底输出安全值
END_CASE

(* —— 段 6：出口单点映射（名实同源，故障码由锁存回放） —— *)
eStateOut := _eState;                    // 状态出口
IF _bFault THEN
    uErrorId := _uFault;                 // 故障锁存码回放（不在故障相按当下输入重推）
ELSE
    uErrorId := _uInfo;                  // 信息码
END_IF
bError := _bFault;                       // 故障出口派生自锁存（非擦除式覆盖）

END_FUNCTION_BLOCK

(* ---- FB_DL_DryingOvenZone.st ---- *)
// =====================================================================
// FB_DL_DryingOvenZone.st
// 烘箱 8 温区串级控温（比例 + 风量前馈 + 速率限幅 + 独立超温联锁）
// Drying oven 8-zone cascade temperature control FB
// 码位: 16#0002_371F ~ 16#0002_3723 (本件独占 5 槽)
// 修改记录: R29 初版 (按 DISPATCH_R29 序 5)
// =====================================================================
FUNCTION_BLOCK FB_DL_DryingOvenZone
VAR_INPUT
    bEnable         : BOOL  := FALSE;   // 使能 / Enable
    bReset          : BOOL  := FALSE;   // 复位 / Reset
    abZoneEnable    : ARRAY[1..8] OF BOOL;      // 8 区独立使能 / Per-zone enable
    afPv_C          : ARRAY[1..8] OF REAL;      // 8 区实测温度 -20~300 ℃ / Zone PV [degC]
    afSp_C          : ARRAY[1..8] OF REAL;      // 8 区设定温度 0~250 ℃ / Zone SP [degC]
    afKp            : ARRAY[1..8] OF REAL;      // 8 区比例增益 0.1~20 %/K / Zone gain [%/K]
    fFanPct         : REAL  := 0.0;     // 循环风量 0~100 % / Fan duty [%]
    fKff            : REAL  := 0.0;     // 风量前馈系数 0~1 %/% / Fan feedforward [%/%]
    fOvertemp_C     : REAL  := 260.0;   // 超温阈值 50~300 ℃ / Overtemperature limit [degC]
    fRateMax_pct_s  : REAL  := 5.0;     // 输出速率上限 >0 %/s / Output slew limit [%/s]
    bFanRun         : BOOL  := FALSE;   // 风机运行反馈 / Fan running
    tCycle          : TIME  := T#100MS; // 周期 T#10MS~T#2S / Cycle [s]
END_VAR
VAR_OUTPUT
    afOut_pct       : ARRAY[1..8] OF REAL;      // 8 区加热输出 0~100 % / Heater output [%]
    bOvertemp       : BOOL;             // 任一区超温（锁存）/ Any zone overtemp, latched
    uOvertempZone   : USINT;            // 首个超温区号 0=无 / First overtemp zone, 0=none
    bReady          : BOOL;             // 全部区进入带内 / All zones in band
    eState          : E_DL_OvenState;   // 状态 / State
    eErr            : UDINT;            // 错误码 / Error code
END_VAR
VAR
    uIdx            : UDINT;            // 区循环下标 / Zone loop index
    uZi             : INT;              // 1..8 数组下标 / Array subscript 1..8
    uZj2            : INT;              // 清零循环第二下标 / Second subscript for zero loops
    fDevK           : REAL;             // 区偏差 K / Zone deviation [K]
    fSpSafe         : REAL;             // 处理后设定（≤0 按 1 ℃）/ Sanitized SP [degC]
    fOutRaw         : REAL;             // 计算原始输出 / Raw computed output [%]
    fStepMax        : REAL;             // 单拍步长 / Max step per cycle [%]
    fStep           : REAL;             // 本拍实际步长 / Actual step this cycle [%]
    tCycleS         : REAL;             // 周期秒值（钳 ≥0.01）/ Cycle in seconds, clamped [s]
    bAllEnabled     : BOOL;             // 是否存在使能区 / Any zone enabled
    bFanBad         : BOOL;             // 风量非有限标记 / Fan duty non-finite flag
    fFanPctSafe     : REAL;             // 处理后风量 / Sanitized fan duty [%]
    bAnyOver        : BOOL;             // 本拍超温探测 / Overtemp detected this cycle
    uFirstOver      : USINT;            // 本拍首个超温区 / First overtemp zone this cycle
    xFirstScan      : BOOL := TRUE;     // 首扫标记 / First-scan flag
END_VAR

// ---------------------------------------------------------------------
// 代码位表（本件独占，勿复用）:
//   16#0002_371F 信息 正常运行
//   16#0002_3720 故障 任一 afPv_C/afSp_C 非有限，或 tCycle 非法
//   16#0002_3721 故障 fOvertemp_C ≤ 0 / fRateMax_pct_s ≤ 0 / 任一 afKp ≤ 0（组态错）
//   16#0002_3722 信息 bFanRun=FALSE → 前馈禁用（fKff 项按 0 计），调节继续
//   16#0002_3723 故障 任一区 afPv_C ≥ fOvertemp_C → 全输出清零、锁存，解除=bReset 且全部 PV < 阈值-5K
// ---------------------------------------------------------------------

// ---- 周期转秒并钳下限 / Cycle to seconds with clamp ----
tCycleS := TIME_TO_REAL(tCycle) / 1000.0;   // 秒值 / Seconds [s]
IF tCycleS < 0.01 THEN
    tCycleS := 0.01;    // 钳 ≥0.01 s 防步长爆炸 / Clamp minimum 10 ms
END_IF

// ---- 单拍步长 / Max step per cycle ----
fStepMax := fRateMax_pct_s * tCycleS;       // %/s × s = % / Step per cycle [%]

// ---- 超温锁存解除路径（必须可达，R28）：bReset 且全部 PV < 阈值-5K 回差 / Reset path with 5K hysteresis ----
IF bOvertemp AND bReset THEN
    bAnyOver := FALSE;          // 回差判据累加器 / Hysteresis accumulator
    FOR uIdx := 1 TO 8 DO
        uZi := UDINT_TO_INT(uIdx);              // 下标转换 / Subscript conversion
        IF afPv_C[uZi] >= (fOvertemp_C - 5.0) THEN
            bAnyOver := TRUE;   // 仍有区未回落 5K / Zone not cooled by 5K
        END_IF
    END_FOR
    IF NOT bAnyOver THEN
        bOvertemp     := FALSE; // 解除锁存 / Release latch
        uOvertempZone := 0;     // 区号清零 / Clear zone number
        eState := E_DL_OvenState.eIdle; // 回空闲 / Back to idle
    END_IF
END_IF

// ---- 非有限与周期合法性闸（故障级）/ Finite and cycle validity gate ----
IF (tCycle = T#0MS) OR (tCycleS > 2.0)
   OR (fFanPct <> fFanPct) OR (ABS(fFanPct) >= 1.0E12)
   OR (fKff <> fKff) OR (ABS(fKff) >= 1.0E12)
   OR (fOvertemp_C <> fOvertemp_C) OR (ABS(fOvertemp_C) >= 1.0E12)
   OR (fRateMax_pct_s <> fRateMax_pct_s) OR (ABS(fRateMax_pct_s) >= 1.0E12) THEN
    bOvertemp     := FALSE;     // 清锁存避免卡死 / Clear latch to avoid deadlock
    uOvertempZone := 0;         // 区号清零 / Clear zone
    FOR uZi := 1 TO 8 DO
        afOut_pct[uZi] := 0.0;  // 全输出清零（安全侧）/ Zero all outputs
    END_FOR
    bReady := FALSE;            // 就绪失效 / Not ready
    eState := E_DL_OvenState.eFault;    // 故障态（本闸不锁存，可自动恢复）/ Fault state
    eErr   := 16#0002_3720;     // 故障码 / Fault code
    RETURN;                     // 本拍结束 / End of cycle
END_IF

// ---- 各区 PV/SP 非有限逐个判界（多 ARRAY 按各自上界逐个判）/ Per-zone finite check ----
FOR uZi := 1 TO 8 DO
    IF (afPv_C[uZi] <> afPv_C[uZi]) OR (ABS(afPv_C[uZi]) >= 1.0E12)
       OR (afSp_C[uZi] <> afSp_C[uZi]) OR (ABS(afSp_C[uZi]) >= 1.0E12) THEN
        FOR uZj2 := 1 TO 8 DO
            afOut_pct[uZj2] := 0.0;  // 全输出清零 / Zero all outputs
        END_FOR
        bReady := FALSE;        // 就绪失效 / Not ready
        eState := E_DL_OvenState.eFault;    // 故障态 / Fault state
        eErr   := 16#0002_3720; // 故障码 / Fault code
        RETURN;                 // 本拍结束 / End of cycle
    END_IF
END_FOR

// ---- 组态错闸 / Configuration fault gate ----
IF (fOvertemp_C <= 0.0) OR (fRateMax_pct_s <= 0.0) THEN
    FOR uZi := 1 TO 8 DO
        afOut_pct[uZi] := 0.0;  // 全输出清零 / Zero all outputs
    END_FOR
    bReady := FALSE;            // 就绪失效 / Not ready
    eState := E_DL_OvenState.eFault;    // 故障态 / Fault state
    eErr   := 16#0002_3721;     // 故障码 / Fault code
    RETURN;                     // 本拍结束 / End of cycle
END_IF
FOR uZi := 1 TO 8 DO
    IF afKp[uZi] <= 0.0 THEN
        FOR uZj2 := 1 TO 8 DO
            afOut_pct[uZj2] := 0.0;  // 全输出清零 / Zero all outputs
        END_FOR
        bReady := FALSE;        // 就绪失效 / Not ready
        eState := E_DL_OvenState.eFault;    // 故障态 / Fault state
        eErr   := 16#0002_3721; // 故障码 / Fault code
        RETURN;                 // 本拍结束 / End of cycle
    END_IF
END_FOR

// ---- 首扫初始化（R16 首扫纪律）/ First-scan initialization ----
IF xFirstScan THEN
    FOR uZi := 1 TO 8 DO
        afOut_pct[uZi] := 0.0;  // 输出从 0 起步 / Outputs start at zero
    END_FOR
    xFirstScan := FALSE;        // 清首扫标记 / Clear flag
END_IF

// ---- 使能撤销：全区输出清零回空闲 / Disable: zero outputs and idle ----
IF NOT bEnable THEN
    FOR uZi := 1 TO 8 DO
        afOut_pct[uZi] := 0.0;  // 全输出清零 / Zero all outputs
    END_FOR
    bReady := FALSE;            // 就绪失效 / Not ready
    eState := E_DL_OvenState.eIdle;     // 空闲态 / Idle state
    eErr   := 16#0002_371F;     // 信息级：空闲正常 / Info: idle normal
    RETURN;                     // 本拍结束 / End of cycle
END_IF

// ---- 使能区存在性检查：全关 → eIdle 输出全 0 / No enabled zone → idle ----
bAllEnabled := FALSE;           // 累加器复位 / Reset accumulator
FOR uZi := 1 TO 8 DO
    IF abZoneEnable[uZi] THEN
        bAllEnabled := TRUE;    // 至少一区使能 / At least one zone enabled
    END_IF
END_FOR
IF NOT bAllEnabled THEN
    FOR uZi := 1 TO 8 DO
        afOut_pct[uZi] := 0.0;  // 全输出清零 / Zero all outputs
    END_FOR
    bReady := FALSE;            // 就绪失效 / Not ready
    eState := E_DL_OvenState.eIdle;     // 空闲态 / Idle state
    eErr   := 16#0002_371F;     // 信息级：空闲正常 / Info: idle normal
    RETURN;                     // 本拍结束 / End of cycle
END_IF

// ---- 风量前馈有效性：bFanRun=FALSE → 前馈项按 0 计 / Feedforward disabled without fan ----
bFanBad := FALSE;               // 标记复位 / Reset flag
fFanPctSafe := fFanPct;         // 原值采用 / Adopt as-is
IF NOT bFanRun THEN
    fFanPctSafe := 0.0;         // 前馈禁用（不是零输出）/ FF disabled, control continues
END_IF

// ---- 超温探测（超温优先于调节）/ Overtemp detection has priority ----
bAnyOver   := FALSE;            // 探测复位 / Reset detection
uFirstOver := 0;                // 首区清零 / Clear first zone
FOR uZi := 1 TO 8 DO
    IF afPv_C[uZi] >= fOvertemp_C THEN
        bAnyOver := TRUE;       // 探测到超温 / Overtemp found
        IF uFirstOver = 0 THEN
            uFirstOver := INT_TO_USINT(uZi);    // 记录首区 / Record first zone
        END_IF
    END_IF
END_FOR

IF bAnyOver THEN
    // 超温路径：全输出清零 + 故障锁存，绝不边降温边加热 / Overtemp: zero all, latch fault
    FOR uZi := 1 TO 8 DO
        afOut_pct[uZi] := 0.0;  // 全输出清零（安全侧）/ Zero all outputs
    END_FOR
    bOvertemp     := TRUE;      // 锁存 / Latch
    uOvertempZone := uFirstOver;    // 记首区 / First zone
    bReady        := FALSE;     // 就绪失效 / Not ready
    eState        := E_DL_OvenState.eFault;     // 故障态 / Fault state
    eErr          := 16#0002_3723;      // 故障码 / Fault code
    RETURN;                     // 本拍结束 / End of cycle
END_IF

// ---- 正常调节路径（eRun）：逐区比例 + 前馈 + 速率限幅 / Normal control path ----
eState := E_DL_OvenState.eRun;      // 运行态 / Run state
bReady := TRUE;                     // 就绪假设成立，区带外再翻 false / Assume ready, clear per zone
FOR uZi := 1 TO 8 DO
    IF abZoneEnable[uZi] THEN
        // 设定 ≤0 按 1 ℃ 处理（防冻结工况斜率无穷）/ SP ≤0 treated as 1 degC
        IF afSp_C[uZi] <= 0.0 THEN
            fSpSafe := 1.0;     // 防斜率无穷 / Guard slope
        ELSE
            fSpSafe := afSp_C[uZi]; // 原值 / As-is
        END_IF
        fDevK := fSpSafe - afPv_C[uZi];     // 偏差 = SP - PV / Deviation [K]
        // 比例项 + 风量前馈项 / Proportional + fan feedforward term
        fOutRaw := afKp[uZi] * fDevK + fKff * fFanPctSafe;  // 原始输出 [%]
        // 前馈禁用信息级（bFanRun=FALSE 且 fKff>0 时提示）/ FF disabled info
        IF (NOT bFanRun) AND (fKff > 0.0) THEN
            eErr := 16#0002_3722;   // 信息级：前馈禁用 / Info: FF disabled
        END_IF
        // 输出限幅 0~100 % / Clamp 0..100
        IF fOutRaw < 0.0 THEN
            fOutRaw := 0.0;     // 下限 / Lower clamp
        ELSIF fOutRaw > 100.0 THEN
            fOutRaw := 100.0;   // 上限 / Upper clamp
        END_IF
        // 速率限幅（单拍增量 ≤ fStepMax）/ Slew limit per cycle
        fStep := fOutRaw - afOut_pct[uZi];  // 期望步长 / Desired step [%]
        IF fStep > fStepMax THEN
            fStep := fStepMax;      // 正向限速 / Positive slew
        ELSIF fStep < -fStepMax THEN
            fStep := -fStepMax;     // 负向限速 / Negative slew
        END_IF
        afOut_pct[uZi] := afOut_pct[uZi] + fStep;   // 采纳步长 / Adopt step
        // 带内判（±2 K 带容差）/ In-band check (±2 K tolerance)
        IF ABS(fSpSafe - afPv_C[uZi]) > 2.0 THEN
            bReady := FALSE;    // 区带外 → 就绪失效 / Zone out of band
        END_IF
    ELSE
        afOut_pct[uZi] := 0.0;  // 禁用区输出保持 0 / Disabled zone output zero
    END_IF
END_FOR

// 未在任何分支改写 eErr 时补正常码 / Default normal code if untouched
IF eErr <> 16#0002_3722 THEN
    eErr := 16#0002_371F;       // 信息级：正常运行 / Info: normal run
END_IF

END_FUNCTION_BLOCK

(* ---- FB_DL_DuctLeakRateEst.st ---- *)
(*
  FB_DL_DuctLeakRateEst  —  风管漏风率估算（流量差法 + 静压修正 + 分级判据） / Duct air-leakage rate estimation by flow difference with static-pressure correction and class grading
  分类 Category : DL_Algo
  版本 Version  : 1.0.0
  来源 Source   : t1-2-oscat-building — 楼宇风管验收算法族深化
  溯源 Origin   : 道莅 clean-room 实现；漏风率 = 100×(送风-回风)/送风 与静压线性修正为公开暖通测试算法，未复制任何源码行
  功能 Function : 1) 流量差法：_fLeakPct = 100 × (fSupplyM3h - fReturnM3h) / fSupplyM3h，
                  分母 <= 1.0E-6 判非法（除零前置守卫）；
                  2) 静压修正：_fCorrPct = (fStaticPa - fStaticRefPa) / 10.0 × fPressCorrPctPer10Pa，
                  修正后 _fLeakCorr = _fLeakPct - _fCorrPct（除数为常量 10.0）；
                  3) 向上取整到 0.1%：先实数上限兜底 → 截断 → 按余量进位（正好整除不 +1，
                  禁 TRUNC(x)+1 写法，R28-2）；
                  4) 分级：A/B/C 三档阈值判据，越 C 档为不合格（eReject）。
                  5) 本件只有故障码、无信息码（派单硬约束）。
  接口 Interface: 输入送/回风量、静压与参考静压、修正系数、三档阈值；输出漏风率/分级/码
  边界 Boundary : ① 组态闸：fSupplyM3h <= 1.0E-6、fPressCorrPctPer10Pa < 0.0、
                  fClassAPct < 0.0 或 fClassBPct <= fClassAPct 或 fClassCPct <= fClassBPct
                  → 0386 锁存；② 送/回风量或静压非有限（NaN 自反 + Inf 差值自减）→ 0386 锁存；
                  ③ 取整前实数上限兜底（2.147483E9 对应 DINT 可表上界），防 LREAL→DINT 溢出；
                  ④ 回风量大于送风量时漏风率为负，按死区归 0（-0.05% 容差带），不判故障；
                  ⑤ 零全局耦合：无 GVL / VAR_EXTERNAL / %I %Q %M 直接地址。
  依赖 Depends  : Standard.library（R_TRIG）
  码表 Error codes（Algo 段 0002，故障窗口 0386；本件无信息码）:
    16#0002_0386 故障级：漏风率估算故障总码（组态非法 / 风量或静压非有限 / 送风量为零导致除零），
                 锁存至 bReset 上升沿；归因见 eCause，不新增码位（派单硬约束单码）
  修订历史 Revision :
    2026-11-19  v1.0.0  R43 首版（批次 2 · 序号 10）
*)

TYPE E_DL_DlrState :
(
    eIdle  := 0,      // 未使能待估算 / Idle, waiting evaluation
    eRun   := 10,     // 估算运行中 / Evaluation active
    eFault := 90      // 故障锁存相 / Fault latched phase
);
END_TYPE

TYPE E_DL_DlrClass :
(
    eNone    := 0,    // 未分级 / Not graded
    eClassA  := 1,    // A 级（最严） / Class A, tightest
    eClassB  := 2,    // B 级 / Class B
    eClassC  := 3,    // C 级 / Class C
    eReject  := 4     // 不合格（越 C 档） / Rejected, beyond class C
);
END_TYPE

TYPE E_DL_DlrCause :
(
    eNone      := 0,  // 无故障成因 / No cause
    eCfgIllegal:= 1,  // 组态非法 / Illegal configuration
    eNonFinite := 2,  // 输入非有限 / Non-finite input
    eDivZero   := 3   // 送风量过小（除零风险） / Supply flow too small
);
END_TYPE

FUNCTION_BLOCK FB_DL_DuctLeakRateEst
VAR_INPUT
    fSupplyM3h        : REAL := 0.0;      // 送风量 [m³/h]，域 > 0 / Supply air flow
    fReturnM3h        : REAL := 0.0;      // 回风量 [m³/h] / Return air flow
    fStaticPa         : REAL := 0.0;      // 实测静压 [Pa] / Measured static pressure
    fStaticRefPa      : REAL := 0.0;      // 参考静压 [Pa] / Reference static pressure
    fPressCorrPctPer10Pa : REAL := 0.5;   // 每 10 Pa 修正百分比 [%/10Pa]，域 >= 0 / Correction per 10 Pa
    fClassAPct        : REAL := 1.0;      // A 级上限 [%] / Class A limit
    fClassBPct        : REAL := 3.0;      // B 级上限 [%] / Class B limit
    fClassCPct        : REAL := 6.0;      // C 级上限 [%] / Class C limit
    fNegDeadbandPct   : REAL := 0.05;     // 负值死区 [%]，域 >= 0 / Negative deadband
    bEnable           : BOOL := FALSE;    // 估算使能（电平）[-] / Evaluation enable
    bReset            : BOOL := FALSE;    // 复位命令，上升沿清故障 [-] / Reset edge
END_VAR
VAR_OUTPUT
    eState            : E_DL_DlrState;    // 状态出口，段 6 单点映射 / State outlet
    eClass            : E_DL_DlrClass;    // 分级出口 / Grading outlet
    eCause            : E_DL_DlrCause;    // 故障成因出口（R190） / Fault cause outlet
    fLeakPct          : REAL;             // 原始漏风率 [%] / Raw leakage rate
    fLeakCorrPct      : REAL;             // 静压修正后漏风率 [%] / Corrected leakage rate
    fLeakCeilPct      : REAL;             // 向上取整到 0.1% 的漏风率 [%] / Ceil to 0.1 %
    bError            : BOOL;             // 故障锁存标志 [-] / Fault latch flag
    nErrId            : UDINT;            // 故障码，0 = 无故障（本件无信息码） / Fault code only
END_VAR
VAR
    _eState           : E_DL_DlrState := E_DL_DlrState.eIdle;     // 内部相位（CASE 唯一写入目标） / Internal phase
    _eClass           : E_DL_DlrClass := E_DL_DlrClass.eNone;     // 分级槽（每拍重算） / Grading slot
    _eCause           : E_DL_DlrCause := E_DL_DlrCause.eNone;     // 故障成因锁存（锁存量） / Latched cause
    rtReset           : R_TRIG;           // 复位沿实例，每周期无条件调用 / Reset edge
    _fDiffM3h         : REAL;             // 送回风量差 [m³/h]（当拍量） / Flow difference
    _fCorrPct         : REAL;             // 静压修正量 [%]（当拍量） / Pressure correction
    _fScaled          : REAL;             // 取整中间量（×10 后） / Scaling intermediate
    _iScaled          : DINT;             // 截断后整数（×10） / Truncated integer
    _bNonFin          : BOOL;             // 输入非有限当拍量 [-] / Non-finite input
    _bDivRisk         : BOOL;             // 除零风险当拍量 [-] / Divide risk
    _bCfgBad          : BOOL;             // 组态非法当拍量 [-] / Config illegal
    _bFault           : BOOL;             // 故障锁存位（锁存量） / Latched fault bit
    _uFault           : UDINT;            // 故障码锁存（锁存量） / Latched fault code
END_VAR

(* —— 段 0：沿实例无条件周期刷新 + 当拍量判据 —— *)
_bNonFin := (fSupplyM3h <> fSupplyM3h) OR (fReturnM3h <> fReturnM3h) OR (fStaticPa <> fStaticPa)
         OR ((fSupplyM3h - fSupplyM3h) <> (fSupplyM3h - fSupplyM3h))
         OR ((fReturnM3h - fReturnM3h) <> (fReturnM3h - fReturnM3h))
         OR ((fStaticPa - fStaticPa) <> (fStaticPa - fStaticPa));            // NaN 自反 + Inf 差值自减 / NaN and Inf detection
_bDivRisk := fSupplyM3h <= 1.0E-6;                                           // 送风量过小（除零风险） / Divide risk
_bCfgBad := _bDivRisk OR (fPressCorrPctPer10Pa < 0.0) OR (fClassAPct < 0.0)
            OR (fClassBPct <= fClassAPct) OR (fClassCPct <= fClassBPct)
            OR (fNegDeadbandPct < 0.0);                                      // 组态非法当拍量 / Config illegal
rtReset(CLK := bReset);                                                      // 复位沿，每拍必调 / Reset edge

(* —— 段 1：单拍量预清零（锁存量不入清单；分级槽每拍重算） —— *)
eClass := E_DL_DlrClass.eNone;      // 分级出口缺省未分级 / Grading default
eCause := _eCause;                  // 成因出口映射（锁存量回放，段 6 复核） / Cause outlet
fLeakPct := 0.0;                    // 原始漏风率缺省 0 / Raw rate default
fLeakCorrPct := 0.0;                // 修正后漏风率缺省 0 / Corrected rate default
fLeakCeilPct := 0.0;                // 取整漏风率缺省 0 / Ceil rate default
nErrId := 16#0000_0000;             // 故障码缺省无故障 / Fault code default

(* —— 段 2：复位沿 + 组态域闸 —— *)
IF rtReset.Q THEN                              // rtReset.Q = 当拍量 / current scan
    _bFault := FALSE;                          // 清故障锁存位（锁存量） / Clear fault latch
    _uFault := 16#0000_0000;                   // 清故障锁存码（锁存量） / Clear fault code
    _eCause := E_DL_DlrCause.eNone;            // 清成因（锁存量） / Clear cause
    IF _eState = E_DL_DlrState.eFault THEN
        _eState := E_DL_DlrState.eIdle;        // 故障相迁出：回未使能 / Fault exit to idle
    END_IF
END_IF
IF _bNonFin THEN                               // 非有限锁存（独立归因） / Non-finite latch
    _uFault := 16#0002_0386;                   // 故障级：估算故障总码 / Algo fault code
    _eCause := E_DL_DlrCause.eNonFinite;       // 归因：非有限 / Cause: non-finite
    _bFault := TRUE;                           // 标志与码位配对（R45） / Flag paired with code
END_IF
IF _bCfgBad THEN                               // 组态域闸 / Config gate
    _uFault := 16#0002_0386;
    IF _bDivRisk THEN
        _eCause := E_DL_DlrCause.eDivZero;     // 归因：除零风险 / Cause: divide risk
    ELSE
        _eCause := E_DL_DlrCause.eCfgIllegal;  // 归因：组态非法 / Cause: illegal config
    END_IF
    _bFault := TRUE;
END_IF

(* —— 段 3：漏风率与分级（仅无故障时计算；除数为已校验正域） —— *)
IF (NOT _bFault) AND (_eState = E_DL_DlrState.eRun) THEN
    _fDiffM3h := fSupplyM3h - fReturnM3h;                          // 流量差 / Flow difference
    fLeakPct := 100.0 * _fDiffM3h / fSupplyM3h;                    // 原始漏风率（分母已守卫） / Raw rate
    _fCorrPct := (fStaticPa - fStaticRefPa) / 10.0 * fPressCorrPctPer10Pa;   // 静压修正（除常量 10.0） / Correction
    fLeakCorrPct := fLeakPct - _fCorrPct;                          // 修正后漏风率 / Corrected rate
    IF (fLeakCorrPct < 0.0) AND (ABS(fLeakCorrPct) <= fNegDeadbandPct) THEN
        fLeakCorrPct := 0.0;                                       // 负值死区归 0 / Negative deadband
    END_IF
    _fScaled := fLeakCorrPct * 10.0;                               // 放大 10 倍进入整数域 / Scale by ten
    IF _fScaled >= 2.147483E9 THEN                                 // 实数上限兜底（DINT 可表上界） / Real upper guard
        _fScaled := 2.147483E9;
    ELSIF _fScaled <= -2.147483E9 THEN                             // 实数下限兜底 / Real lower guard
        _fScaled := -2.147483E9;
    END_IF
    _iScaled := LREAL_TO_DINT(LREAL(_fScaled));                    // 截断取整 / Truncate
    IF LREAL(_iScaled) < LREAL(_fScaled) - 1.0E-9 THEN             // 余量进位（正好整除不进位） / Ceiling by remainder
        _iScaled := _iScaled + 1;
    END_IF
    fLeakCeilPct := DINT_TO_REAL(_iScaled) * 0.1;                  // 还原为 0.1% 步长 / Restore 0.1 % step
    IF fLeakCeilPct <= fClassAPct THEN
        _eClass := E_DL_DlrClass.eClassA;                          // A 级 / Class A
    ELSIF fLeakCeilPct <= fClassBPct THEN
        _eClass := E_DL_DlrClass.eClassB;                          // B 级 / Class B
    ELSIF fLeakCeilPct <= fClassCPct THEN
        _eClass := E_DL_DlrClass.eClassC;                          // C 级 / Class C
    ELSE
        _eClass := E_DL_DlrClass.eReject;                          // 不合格（ELSE 兜底） / Rejected fallback
    END_IF
END_IF

(* —— 段 4：故障解除式（R240；全当拍量）：rtReset.Q / NOT _bNonFin / NOT _bCfgBad —— *)
IF rtReset.Q AND (NOT _bNonFin) AND (NOT _bCfgBad) THEN
    _bFault := FALSE;                          // 清故障锁存位（锁存量） / Clear fault latch
    _uFault := 16#0000_0000;                   // 清故障锁存码（锁存量） / Clear fault code
    _eCause := E_DL_DlrCause.eNone;            // 清成因（锁存量） / Clear cause
END_IF

(* —— 段 4A：故障锁存相位迁移闸 —— *)
IF _bFault AND (_eState <> E_DL_DlrState.eFault) THEN
    _eState := E_DL_DlrState.eFault;           // 锁存即入故障相 / Latch enters fault phase
END_IF

(* —— 段 5：相位机（CASE 全覆盖 + ELSE 兜底） —— *)
CASE _eState OF

E_DL_DlrState.eIdle:
    IF bEnable AND (NOT _bFault) THEN          // 使能条件 / Enable gate
        _eState := E_DL_DlrState.eRun;         // 进估算相 / Enter evaluation
    END_IF

E_DL_DlrState.eRun:
    IF NOT bEnable THEN                        // 撤使能：回未使能（前置消失） / Disable returns idle
        _eState := E_DL_DlrState.eIdle;
    END_IF

E_DL_DlrState.eFault:
    ;                                          // 故障相：仅段 4 复位沿可迁出 / Only reset exits

ELSE
    _uFault := 16#0002_0386;                   // 故障级：非法相位兜底（归并总码） / Illegal phase fallback
    _eCause := E_DL_DlrCause.eCfgIllegal;      // 归因：相位非法归并组态 / Cause: phase illegal
    _bFault := TRUE;
    _eState := E_DL_DlrState.eFault;           // 强制回故障相 / Force fault phase

END_CASE

(* —— 段 6：出口单点映射（名实同源；锁存码回放，禁同拍抹除） —— *)
IF _bFault THEN
    nErrId := _uFault;                         // 故障锁存码回放 / Replay latched code
    eClass := E_DL_DlrClass.eNone;             // 故障相分级强制未分级 / Grading forced none
    fLeakCeilPct := 0.0;                       // 故障相取整值强制 0（安全侧） / Ceil forced zero
ELSE
    nErrId := 16#0000_0000;                    // 无故障：本件无信息码 / No fault, no info code
    eClass := _eClass;                         // 分级出口 / Grading outlet
END_IF
bError := _bFault;                             // 故障标志同源 / Flag from latch
eState := _eState;                             // 状态出口 / State outlet
eCause := _eCause;                             // 成因出口 / Cause outlet

END_FUNCTION_BLOCK

(* ---- FB_DL_DuctStaticReset.st ---- *)
//==============================================================================
// 功能块：FB_DL_DuctStaticReset ｜ 中文名称：风管静压设定重置
// 所属子库：DL_Algo ｜ 版本：v1.0.0 ｜ 兼容：CODESYS V3.5+ / TwinCAT 3 / 汇川 InoProShop
// 功能描述：风管静压设定重置（TSP 修剪侧单件）：最不利末端阀位落在目
//           标带 [100−band, 100) 视为合适（带内保持）；阀位顶满 100%
//           （超带）→ 设定按增益上抬；阀位低于带下沿 → 设定按增益下
//           调。设定变化经斜率限制（fRatePaPerS，由 uDeltaTimeMs 显式
//           积分，禁系统时间函数），上下限钳位。阀位反馈无效（bFbValid
//           为假）→ 保持上次设定并发 3502（信息级，不置 bError）；设
//           定已顶上限而阀位仍满开 → 3501 能力不足，不再继续抬设定。
//           只算设定值，不控变频器（风机调速由上位裁决，本件零执行输
//           出）。规格 §4.8 引脚表未给反馈有效性输入、但其边界行为③
//           与输出表均要求 bFbInvalid/3502 语义，故增补 VAR_INPUT
//           bFbValid（默认 TRUE）承载上游质量位（主动偏离披露，见修
//           订历史）。
// 开源溯源 (Origin)：道莅原创实现（参考 公开工程惯例 分类与参数域）
// 单位表：阀位[百分数] / 静压[Pa] / 目标带[百分数] / 增益[Pa每百分数] / 斜率[Pa每s] / 扫描间隔[ms]
// 错误码表：16#0002_3501 信息级（静压设定已顶上限且阀位仍全开，风机能
//           力不足，不再抬设定，不置 bError）/ 16#0002_3502 信息级（阀
//           位反馈无效，保持上次设定，不置 bError）/ 16#0002_3505 预留
//           禁用（不得挪用）/ 16#0002_3510 故障级（静压上下限倒置或
//           算法组态非法（带宽/增益/斜率非正），置 bError）/
//           16#0002_3511 故障级（输入非有限，置 bError，设定回下限安
//           全侧防过压）/ 16#0002_3512 预留禁用（不得挪用）
// 状态机：E_DL_DuctStaticState（eIdle=0 / eInBand=10 / eAdjustUp=20 /
//           eAdjustDown=30 / eFbHold=40 / eFault=99），CASE 含 ELSE 兜
//           底，ELSE 复用 3511（§3 未为本件单列兜底槽，不得越段加码）
//           并回下限安全侧
// 边界行为：① fStaticMinPa 大于等于 fStaticMaxPa 或带宽/增益/斜率非正
//           → 故障 3510；② 阀位域钳 0~100（轻域外按边界值照算）；
//           ③ 阀位反馈无效（bFbValid 为假）→ 保持上次设定 + 信息 3502，
//           挂 eFbHold 相，退出条件两条：反馈恢复（按带位回归工作相）
//           或失能（回待机）；④ 设定已达上限而阀位仍 100% → 信息 3501
//           + bAtLimit，不再继续抬设定；⑤ 斜率限制用 uDeltaTimeMs 显
//           式积分（LREAL 中间量，禁系统时间函数），uDeltaTimeMs 为 0
//           时本拍不动；⑥ 非有限（NaN 自反判 + Inf 幅值上限判，R79）
//           → 故障 3511，设定回 fStaticMinPa 安全侧（防过压）；⑦ 失
//           能 → 保持设定（静压突变会导致末端振荡）+ bValid := FALSE；
//           ⑧ 带语义披露：阀位落在 [100−band, 100) 带内保持，阀位 =
//           100% 视为顶带超限（需上抬），与验收向量 ①② 口径一致；
//           ⑨ 首拍设定从下限起坡（首拍不出未知值）。
// 修订历史：v1.0.0 2026-11-17 首版（R25 派单 · §4.8）
//==============================================================================
(*------------------------------------------------------------------------------
 * 枚举: E_DL_DuctStaticState（归属 DL_Algo，与 FB_DL_DuctStaticReset 同文件）
 *----------------------------------------------------------------------------*)
TYPE E_DL_DuctStaticState :
(
    eIdle       := 0,   // 失能/待机：设定保持，静压不突变 / Idle: setpoint held, no static jump
    eInBand     := 10,  // 阀位带内：设定保持 / In-band: damper within target band, setpoint held
    eAdjustUp   := 20,  // 阀位顶带：设定按斜率上抬 / Damper at band top: setpoint raised by rate
    eAdjustDown := 30,  // 阀位低于带：设定按斜率下调 / Damper below band: setpoint lowered by rate
    eFbHold     := 40,  // 反馈无效保持：设定保持，等反馈恢复 / Feedback-invalid hold: setpoint held
    eFault      := 99   // 故障兜底态：组态非法/非有限/非法状态，设定回下限 / Fault fallback, setpoint at floor
);
END_TYPE
FUNCTION_BLOCK FB_DL_DuctStaticReset
VAR_INPUT
    fWorstDamperPct : LREAL;                   // 最不利末端阀位 [百分数] / Worst-zone damper position [percent]
    fStaticMinPa  : LREAL;                     // 静压设定下限 [Pa] / Static setpoint floor [Pa]
    fStaticMaxPa  : LREAL;                     // 静压设定上限 [Pa] / Static setpoint ceiling [Pa]
    fBandPct      : LREAL := 10.0;             // 阀位目标带 [百分数]，带 = [100−band, 100) / Damper target band [percent]
    fGainPaPerPct : LREAL := 2.0;              // 增益 [Pa每百分数] / Gain [Pa per percent]
    fRatePaPerS   : LREAL := 5.0;              // 设定斜率 [Pa每s] / Setpoint rate limit [Pa per s]
    bFbValid      : BOOL := TRUE;              // 阀位反馈有效性质量位（规格补遗引脚，见修订历史）/ Damper feedback validity, spec-gap pin
    uDeltaTimeMs  : UDINT;                     // 扫描间隔 [ms]，调用方注入，禁用系统时间函数 / Scan interval [ms], caller-injected
    bEnable       : BOOL;                      // 总使能 / Master enable
    bReset        : BOOL;                      // 复位，上升沿清状态与设定 / Reset, rising edge clears state and setpoint
END_VAR
VAR_OUTPUT
    fStaticSetPa  : LREAL;                     // 静压设定 [Pa]，失能保持 / Static setpoint [Pa], held on disable
    bAtLimit      : BOOL;                      // 设定顶上限且阀位仍全开，能力不足 / Setpoint at ceiling with damper full open
    fErrPct       : LREAL;                     // 带偏差 [百分数]，阀位减带下沿，负 = 低于带 / Band deviation [percent], damper minus band floor
    bFbInvalid    : BOOL;                      // 阀位反馈无效标志 / Damper feedback invalid flag
    eErr          : UDINT;                     // 错误码，0 = 无错，码位 16#0002_3501 起信息级、16#0002_3510 起故障级（分带见错误码表） / Error code, 0 = no error, band info/fault per the code table
    bError        : BOOL;                      // 故障级标志，仅故障级错误置位 / Fault-class flag, set only on fault-level codes
    bValid        : BOOL;                      // 设定数据可用标志，失能/故障闸显式 FALSE / Setpoint usable flag, explicit FALSE on disable/fault gates
    eState        : E_DL_DuctStaticState;      // 主状态机当前状态 / Current state of the main state machine
END_VAR
VAR
    fbReset       : R_TRIG;                    // 复位上升沿检测实例 / Reset rising edge detector
    fDamperClamped : LREAL;                    // 钳位后阀位 [百分数] / Clamped damper position [percent]
    fBandFloor    : LREAL;                     // 带下沿 [百分数] / Band floor [percent]
    fStepPa       : LREAL;                     // 本拍允许步长 [Pa]（斜率乘时长）/ Allowed step this scan [Pa]
    fDeltaPa      : LREAL;                     // 本拍目标增量 [Pa]（增益乘带偏差）/ Target delta this scan [Pa]
    fDeltaApplied : LREAL;                     // 本拍实际增量 [Pa]（步长限幅后）/ Applied delta after rate limit [Pa]
    fSetTarget    : LREAL;                     // 限幅前目标设定 [Pa] / Pre-limit target setpoint [Pa]
    bFirstScan    : BOOL := TRUE;              // 首拍初始化标志 / First-scan initialization flag
END_VAR
VAR CONSTANT
    DL_DSR_CODE_INFO_1 : UDINT := 16#0002_3501;   // 信息级槽 1（顶上限且阀位全开） / info slot 1
    DL_DSR_CODE_INFO_2 : UDINT := 16#0002_3502;   // 信息级槽 2（反馈无效保持设定） / info slot 2
    DL_DSR_CODE_RSV_1  : UDINT := 16#0002_3505;   // 预留禁用（不得挪用） / reserved, do not use
    DL_DSR_CODE_FLT_1  : UDINT := 16#0002_3510;   // 故障级槽 1（静压界倒置或组态非法） / fault slot 1
    DL_DSR_CODE_FLT_2  : UDINT := 16#0002_3511;   // 故障级槽 2（输入非有限） / fault slot 2
    DL_DSR_CODE_RSV_2  : UDINT := 16#0002_3512;   // 预留禁用（不得挪用） / reserved, do not use
    DL_DS_ZERO    : LREAL := 0.0;              // 零值常量，避免裸字面量 [—] / Zero constant, avoids a bare literal
    DL_DS_TOL     : LREAL := 1.0E-6;           // 浮点比较容差 [—] / Float comparison tolerance
    DL_DS_INF     : LREAL := 1.7976931348623157E308;  // LREAL 幅值上限，Inf 判据 / LREAL magnitude ceiling, Inf criterion
    DL_DS_PCT_MAX : LREAL := 100.0;            // 阀位域上限 [百分数] / Damper domain ceiling [percent]
    DL_DS_MS_PER_S : LREAL := 1000.0;          // 毫秒转秒系数 [s/ms] / Ms-to-s factor
END_VAR

(*------------------------------------------------------------------------------
 * 段 1｜无条件刷新区（红线 5）：复位沿检测在任何分支之外周期调用
 *----------------------------------------------------------------------------*)
fbReset(CLK := bReset);                        // 复位沿检测无条件刷新 / reset edge refreshed unconditionally

(*------------------------------------------------------------------------------
 * 段 2｜复位沿处理（改写置于沿后，防吞沿 R39）
 *----------------------------------------------------------------------------*)
IF fbReset.Q THEN
    eState  := E_DL_DuctStaticState.eIdle;
    eErr    := 16#0000_0000;                   // 复位清码 / reset clears code
    bError  := FALSE;                          // 复位清故障 / reset clears fault
    bAtLimit := FALSE;                         // 贴限标志清 / at-limit flag cleared
    bFbInvalid := FALSE;                       // 反馈无效标志清 / invalid flag cleared
    bFirstScan := TRUE;                        // 重新首拍化 / re-initialize first scan
    fStaticSetPa := DL_DS_ZERO;                // 设定清零待首拍初始化 / setpoint zeroed, awaits first-scan init
END_IF

(*------------------------------------------------------------------------------
 * 段 3｜非有限输入闸（浮点引脚逐个：NaN 自反判 + Inf 幅值上限判，R79）
 *       命中即设定回下限安全侧（防过压）
 *----------------------------------------------------------------------------*)
IF (fWorstDamperPct <> fWorstDamperPct) OR (ABS(fWorstDamperPct) >= DL_DS_INF)
   OR (fStaticMinPa <> fStaticMinPa) OR (ABS(fStaticMinPa) >= DL_DS_INF)
   OR (fStaticMaxPa <> fStaticMaxPa) OR (ABS(fStaticMaxPa) >= DL_DS_INF)
   OR (fBandPct <> fBandPct) OR (ABS(fBandPct) >= DL_DS_INF)
   OR (fGainPaPerPct <> fGainPaPerPct) OR (ABS(fGainPaPerPct) >= DL_DS_INF)
   OR (fRatePaPerS <> fRatePaPerS) OR (ABS(fRatePaPerS) >= DL_DS_INF) THEN
    eState       := E_DL_DuctStaticState.eFault;
    eErr         := DL_DSR_CODE_FLT_2;             // 故障级：输入非有限 / fault: non-finite input
    bError       := TRUE;                      // 故障级必置 bError（R45 配对）/ fault-class pairs with bError
    bValid       := FALSE;                     // 输出不可用 / outputs unusable
    fStaticSetPa := fStaticMinPa;              // 设定回下限安全侧（防过压）/ setpoint to floor, safe side against overpressure
    bAtLimit := FALSE;                         // 故障态不判贴限 / at-limit not judged in fault
    bFbInvalid := FALSE;                       // 故障态不判反馈无效 / invalid not judged in fault
    fErrPct := DL_DS_ZERO;                     // 带偏差出口清零 / band deviation zeroed
    RETURN;
END_IF

(*------------------------------------------------------------------------------
 * 段 4｜组态合法性闸（静压界倒置/带宽/增益/斜率非正）
 *----------------------------------------------------------------------------*)
IF (fStaticMinPa >= fStaticMaxPa) OR (fBandPct <= DL_DS_TOL)
   OR (fGainPaPerPct <= DL_DS_TOL) OR (fRatePaPerS <= DL_DS_TOL) THEN
    eState       := E_DL_DuctStaticState.eFault;
    eErr         := DL_DSR_CODE_FLT_1;             // 故障级：静压上下限倒置或组态非法 / fault: static band inverted or config invalid
    bError       := TRUE;                      // 故障级必置 bError（R45 配对）/ fault-class pairs with bError
    bValid       := FALSE;                     // 输出不可用 / outputs unusable
    fStaticSetPa := fStaticMinPa;              // 设定回下限安全侧（防过压）/ setpoint to floor, safe side
    bAtLimit := FALSE;                         // 故障态不判贴限 / at-limit not judged in fault
    bFbInvalid := FALSE;                       // 故障态不判反馈无效 / invalid not judged in fault
    fErrPct := DL_DS_ZERO;                     // 带偏差出口清零 / band deviation zeroed
    RETURN;
END_IF

(*------------------------------------------------------------------------------
 * 段 5｜首拍初始化：设定从下限起坡（首拍不出未知值）
 *----------------------------------------------------------------------------*)
IF bFirstScan THEN
    fStaticSetPa := fStaticMinPa;              // 首拍设定 = 下限 / first-scan setpoint = floor
    bFirstScan := FALSE;                       // 初始化完成 / initialization done
END_IF

(*------------------------------------------------------------------------------
 * 段 6｜阀位钳位与带偏差计算（域钳 0~100，带下沿 = 100 − band）
 *----------------------------------------------------------------------------*)
fDamperClamped := fWorstDamperPct;             // 阀位工作副本 / working copy
IF fDamperClamped < DL_DS_ZERO THEN
    fDamperClamped := DL_DS_ZERO;              // 低于 0 钳入 / below zero clamped
END_IF
IF fDamperClamped > DL_DS_PCT_MAX THEN
    fDamperClamped := DL_DS_PCT_MAX;           // 高于 100 钳入 / above 100 clamped
END_IF
fBandFloor := DL_DS_PCT_MAX - fBandPct;        // 带下沿 = 100 − band [百分数] / band floor
fErrPct := fDamperClamped - fBandFloor;        // 带偏差：负 = 低于带，0~band = 带内，band = 顶带 / band deviation

(*------------------------------------------------------------------------------
 * 段 7｜状态机：CASE 含 ELSE 兜底（非法状态 → 复用 3511 + 回下限，安全侧）
 *----------------------------------------------------------------------------*)
CASE eState OF

    E_DL_DuctStaticState.eIdle:
        bValid := FALSE;                       // 失能闸显式不可用（R72）/ explicit FALSE on disable gate
        bAtLimit := FALSE;                     // 贴限标志清 / at-limit flag cleared
        bFbInvalid := FALSE;                   // 失能不判反馈无效 / invalid not judged in idle
        eErr := 16#0000_0000;                  // 待机无错 / no error in idle
        bError := FALSE;                       // 待机无故障 / no fault in idle
        IF bEnable THEN
            IF bFbValid THEN
                eState := E_DL_DuctStaticState.eInBand;        // 反馈有效进带内相 / valid feedback enters in-band
            ELSE
                eState := E_DL_DuctStaticState.eFbHold;        // 反馈无效进保持相 / invalid feedback enters hold
            END_IF
        END_IF

    E_DL_DuctStaticState.eInBand:
        bValid := TRUE;                        // 带内设定可用 / setpoint usable in band
        bAtLimit := FALSE;                     // 带内不判贴限 / at-limit not judged in band
        bFbInvalid := FALSE;                   // 反馈有效 / feedback valid
        eErr := 16#0000_0000;                  // 带内无错 / no error in band
        bError := FALSE;                       // 带内无故障 / no fault in band
        IF NOT bEnable THEN
            eState := E_DL_DuctStaticState.eIdle;      // 失能回待机（设定保持）/ disable returns to idle, setpoint held
            bValid := FALSE;                   // 失能闸显式不可用 / explicit FALSE on disable gate
        ELSIF NOT bFbValid THEN
            eState := E_DL_DuctStaticState.eFbHold;    // 反馈无效转保持相 / invalid feedback to hold phase
        ELSIF fErrPct >= fBandPct - DL_DS_TOL THEN     // 阀位顶满 100%（fErrPct 达 band 上沿即阀位 = 100）
            eState := E_DL_DuctStaticState.eAdjustUp;  // 顶带超限转上调相 / at band top enters adjust-up
        ELSIF fErrPct < -DL_DS_TOL THEN                // 阀位低于带下沿
            eState := E_DL_DuctStaticState.eAdjustDown;        // 低于带转下调相 / below band enters adjust-down
        END_IF

    E_DL_DuctStaticState.eAdjustUp:
        bValid := TRUE;                        // 上调相设定可用 / setpoint usable in adjust-up
        bFbInvalid := FALSE;                   // 反馈有效 / feedback valid
        IF NOT bEnable THEN
            eState := E_DL_DuctStaticState.eIdle;
            bValid := FALSE;                   // 失能闸显式不可用 / explicit FALSE on disable gate
        ELSIF NOT bFbValid THEN
            eState := E_DL_DuctStaticState.eFbHold;    // 反馈无效转保持相 / invalid feedback to hold phase
        ELSE
            fStepPa := fRatePaPerS * UDINT_TO_LREAL(uDeltaTimeMs) / DL_DS_MS_PER_S;  // 本拍步长 = 斜率乘时长 [Pa]，间隔 0 即不动 / step = rate times interval
            fDeltaPa := fGainPaPerPct * fErrPct;       // 目标增量 = 增益乘带偏差 [Pa] / target delta = gain times deviation
            IF fDeltaPa > fStepPa THEN
                fDeltaApplied := fStepPa;      // 斜率限幅 / rate-limited
            ELSE
                fDeltaApplied := fDeltaPa;     // 未触斜率 / within rate
            END_IF
            fSetTarget := fStaticSetPa + fDeltaApplied;        // 限幅前目标 [Pa] / pre-limit target
            IF fSetTarget >= fStaticMaxPa - DL_DS_TOL THEN
                fStaticSetPa := fStaticMaxPa;  // 钳到上限 / clamped to ceiling
                IF fDamperClamped >= DL_DS_PCT_MAX - DL_DS_TOL THEN
                    bAtLimit := TRUE;          // 设定顶上限且阀位仍全开：能力不足 / at ceiling with full-open damper
                    eErr := DL_DSR_CODE_INFO_1;        // 信息级：能力不足，不再抬设定 / info: capacity insufficient
                    bError := FALSE;           // 信息级不置 bError / info never raises bError
                ELSE
                    bAtLimit := FALSE;         // 阀位未满开，仅钳位 / damper not full, clamp only
                    eErr := 16#0000_0000;      // 清码 / clear code
                END_IF
            ELSE
                fStaticSetPa := fSetTarget;    // 未触上限照算 / below ceiling, apply
                bAtLimit := FALSE;             // 未贴限 / not at limit
                eErr := 16#0000_0000;          // 清码 / clear code
            END_IF
            IF fErrPct < fBandPct - DL_DS_TOL THEN     // 阀位离开顶带（需求消失退出）/ damper left band top
                IF fErrPct >= -DL_DS_TOL THEN
                    eState := E_DL_DuctStaticState.eInBand;    // 回带内相 / back to in-band
                ELSE
                    eState := E_DL_DuctStaticState.eAdjustDown;        // 落到带下方向 / fell below band
                END_IF
            END_IF
        END_IF

    E_DL_DuctStaticState.eAdjustDown:
        bValid := TRUE;                        // 下调相设定可用 / setpoint usable in adjust-down
        bAtLimit := FALSE;                     // 下调相不判贴限 / at-limit not judged in adjust-down
        bFbInvalid := FALSE;                   // 反馈有效 / feedback valid
        IF NOT bEnable THEN
            eState := E_DL_DuctStaticState.eIdle;
            bValid := FALSE;                   // 失能闸显式不可用 / explicit FALSE on disable gate
        ELSIF NOT bFbValid THEN
            eState := E_DL_DuctStaticState.eFbHold;    // 反馈无效转保持相 / invalid feedback to hold phase
        ELSE
            fStepPa := fRatePaPerS * UDINT_TO_LREAL(uDeltaTimeMs) / DL_DS_MS_PER_S;  // 本拍步长 [Pa] / step this scan
            fDeltaPa := fGainPaPerPct * (DL_DS_ZERO - fErrPct);        // 目标减量 = 增益乘带偏差绝对值 [Pa] / target decrement
            IF fDeltaPa > fStepPa THEN
                fDeltaApplied := fStepPa;      // 斜率限幅 / rate-limited
            ELSE
                fDeltaApplied := fDeltaPa;     // 未触斜率 / within rate
            END_IF
            fSetTarget := fStaticSetPa - fDeltaApplied;        // 限幅前目标 [Pa] / pre-limit target
            IF fSetTarget <= fStaticMinPa + DL_DS_TOL THEN
                fStaticSetPa := fStaticMinPa;  // 钳到下限 / clamped to floor
                eErr := 16#0000_0000;          // 清码 / clear code
            ELSE
                fStaticSetPa := fSetTarget;    // 未触下限照算 / above floor, apply
                eErr := 16#0000_0000;          // 清码 / clear code
            END_IF
            IF (fErrPct >= -DL_DS_TOL) AND (fErrPct < fBandPct - DL_DS_TOL) THEN
                eState := E_DL_DuctStaticState.eInBand;        // 回带相（需求消失退出）/ back to in-band when need gone
            END_IF
        END_IF

    E_DL_DuctStaticState.eFbHold:
        bValid := TRUE;                        // 保持相设定输出仍可用（保持值）/ usable in hold (held setpoint)
        bAtLimit := FALSE;                     // 保持相不判贴限 / at-limit not judged in hold
        bFbInvalid := TRUE;                    // 反馈无效标志保持 / invalid flag held
        eErr := DL_DSR_CODE_INFO_2;            // 信息级：反馈无效保持上次设定 / info: invalid feedback, setpoint held
        bError := FALSE;                       // 信息级不置 bError / info never raises bError
        IF NOT bEnable THEN
            eState := E_DL_DuctStaticState.eIdle;      // 失能回待机（第二条退出条件）/ disable returns to idle, second exit
            bValid := FALSE;                   // 失能闸显式不可用 / explicit FALSE on disable gate
            bFbInvalid := FALSE;               // 失能清标志 / flag cleared on disable
        ELSIF bFbValid THEN
            bFbInvalid := FALSE;               // 反馈恢复（第一条退出条件）/ feedback recovered, first exit
            IF fErrPct >= fBandPct - DL_DS_TOL THEN
                eState := E_DL_DuctStaticState.eAdjustUp;      // 按带位回归上调相 / re-enter by band position
            ELSIF fErrPct < -DL_DS_TOL THEN
                eState := E_DL_DuctStaticState.eAdjustDown;    // 按带位回归下调相 / re-enter by band position
            ELSE
                eState := E_DL_DuctStaticState.eInBand;        // 按带位回归带内相 / re-enter by band position
            END_IF
        END_IF

    ELSE
        eState := E_DL_DuctStaticState.eFault; // 非法状态兜底 / illegal-state fallback
        eErr := DL_DSR_CODE_FLT_2;                 // 兜底复用故障级槽 2（§3 未单列兜底槽，不得越段加码）/ fallback reuses fault slot 2
        bError := TRUE;                        // 故障级必置 bError / fault-class pairs with bError
        bValid := FALSE;                       // 输出不可用 / outputs unusable
        fStaticSetPa := fStaticMinPa;          // 设定回下限安全侧（防过压）/ setpoint to floor, safe side
        bAtLimit := FALSE;                     // 贴限标志清 / at-limit flag cleared
        bFbInvalid := FALSE;                   // 标志清 / flag cleared
END_CASE
END_FUNCTION_BLOCK
